(* IEC 61131-3 sources: daoli-st-library/DL_Algo (part 4) *)

(* ---- FC_DL_AccumulationZoneFillCalc.st ---- *)
(*
  DL Factory R83 | FC_DL_AccumulationZoneFillCalc
  功能：按积放区长度与料箱节距算容量件数，并算当前占位率与满料判定。
  开源溯源：无（clean-room 自研，依据公开工艺公式，来源=行业通用公式，许可证=MIT，借鉴点=公式结构）
  规则：R1-R21 全遵守
*)
FUNCTION FC_DL_AccumulationZoneFillCalc : REAL
VAR_INPUT
    fZoneLenM : REAL; // 积放区有效长度 [m] / Accumulation zone effective length [m]
    fToteLenM : REAL; // 料箱长度 [m] / Tote length [m]
    fGapMinM  : REAL; // 最小净间距 [m] / Minimum clear gap [m]
    iToteCnt  : INT;  // 区内实际料箱数 [件] / Actual totes in zone [-]
END_VAR
VAR_OUTPUT
    iCapCnt : INT;  // 区内理论容量件数 [件] / Theoretical capacity [pcs]
    fOccPct : REAL; // 占位率（实际/容量）[%] / Occupancy ratio [%]
    xFull   : BOOL; // 满料判定（占位率不低于 90%）/ Full flag, occupancy at or above 90 percent
    xValid  : BOOL; // 计算有效性标志 / Calculation validity flag
END_VAR
VAR
    fPitchM : REAL; // 单箱占用节距（箱长+净距）[m] / Per-tote pitch [m]
END_VAR
// 出口预置：四出口统一预置，满料标志预置 FALSE（安全侧）
iCapCnt := 0; fOccPct := 0.0; xFull := FALSE; xValid := FALSE;
// 非有限拦截 + 量纲自检 + 计数器域闸（R20/R21）
IF NOT (fZoneLenM > -1.0E30 AND fZoneLenM < 1.0E30) OR NOT (fToteLenM > -1.0E30 AND fToteLenM < 1.0E30) OR NOT (fGapMinM > -1.0E30 AND fGapMinM < 1.0E30) OR fZoneLenM <= 0.0 OR fToteLenM <= 0.0 OR fGapMinM < 0.0 OR iToteCnt < 0 THEN
    FC_DL_AccumulationZoneFillCalc := -1.0; RETURN; // 哨兵 -1：非有限或量纲/计数越界 / Sentinel -1
END_IF
// 单箱节距：箱长 + 最小净距，同量纲相加得 m
fPitchM := fToteLenM + fGapMinM;    // 单箱节距 [m] / Per-tote pitch [m]
// 容量：区长 ÷ 节距 向下取整（禁 TRUNC+1 写法，R28）；节距分母显式零闸（R4/R21）
IF ABS(fPitchM) > 1.0E-9 THEN       // 节距分母显式零闸 / Explicit zero gate on pitch
    iCapCnt := REAL_TO_INT(fZoneLenM / fPitchM);  // 理论容量 [件] / Theoretical capacity
ELSE
    iCapCnt := 0;                   // 除零防御缺省 [件] / Divide-by-zero default
END_IF
// 占位率：实际 ÷ 容量 × 100，容量为零时按零并标记无效（R4/R21）
IF iCapCnt > 0 THEN
    fOccPct := (INT_TO_REAL(iToteCnt) / INT_TO_REAL(iCapCnt)) * 100.0; // 占位率 [%] / Occupancy [%]
    xValid  := TRUE;                // 链路有效 / Chain valid
ELSE
    fOccPct := 0.0;                 // 容量为零不可算占位率 / Zero capacity, occupancy undefined
    xValid  := FALSE;               // 标记无效 / Flag invalid
END_IF
// 满料判定：占位率不低于 90%（含实际数超过理论容量的挤压工况）
xFull := fOccPct >= 90.0;           // 满料布尔 / Full boolean
FC_DL_AccumulationZoneFillCalc := fOccPct; // 返回占位率 [%] / Return occupancy [%]
END_FUNCTION

(* ---- FC_DL_AirDensity.st ---- *)
(*==============================================================================
 * 组件名称 (Component)  : FC_DL_AirDensity
 * 所属子库 (Sublibrary) : DL_Algo
 * 当前版本 (Version)    : 1.0.0
 * 组件分类 (Category)   : 函数（FUNCTION）· 纯函数 · 湿空气物性（密度）
 * 兼容性   (Platform)   : CODESYS 3.5 / TwinCAT 3 / 汇川 InoProShop / Schneider
 *                         Machine Expert；仅用标准 EXP / ABS / LIMIT
 * 功能描述 (Function)   : 按干空气与水蒸气分压叠加法计算湿空气密度
 *                         密度 = 干空气分压 除以 (干空气气体常数 乘以 绝对温度)
 *                                + 水蒸气分压 除以 (水蒸气气体常数 乘以 绝对温度)
 *                         单位为千克每立方米。饱和蒸汽压用 Magnus-Tetens 式计算。
 *                         用于风量质量流量换算（风机功率核算、风管风速换算）、
 *                         洁净室换气次数、烘干与涂布风量配比、空压站产气量折算。
 * 与既有件边界 (Boundary): FC_DL_HumidAirEnthalpy 出比焓（焦耳每克）；
 *                         FC_DL_DewPointCalc 出露点（摄氏度）；本件出密度
 *                         （千克每立方米）。三件共享同一 Magnus 常量口径，
 *                         但各自内联实现，禁止互相调用（泳道内零依赖），
 *                         保证任一件单独移植时不需要再带两个依赖件。
 * 精度声明 (Accuracy)   : 在零下 10 度到 50 度域内，相对误差小于 0.5 个百分点
 *                         （公开文献口径）；超出该域仅供趋势参考。这是本库对
 *                         OSCAT 同类函数行为定义的收窄，按 R11 留档。
 * 设计要点 (Key notes)  : ① 干空气分压必须防负：高湿低压的极端组态会出现
 *                           水蒸气分压大于总压，物理上不可能，但组态可给出；
 *                           出现即钳到 0 并置码，绝不输出负密度；
 *                         ② Magnus 式分母（243.12 加温度）在零下 40 度时为
 *                           203.12，恒大于 0，温度下限已保证无除零；
 *                         ③ 绝对温度由温度下限保证不小于 233.15 开，恒正；
 *                         ④ 域校验采用「钳位后继续算」策略：现场宁可要一个
 *                           标注为近似的密度值，也不要因为传感器越量程就断链。
 * 开源溯源 (Origin)     : oscat-building。参考 OSCAT 公开函数库 Building 分类
 *                         中空气密度函数的功能分类与参数域（温度 / 压力 /
 *                         湿度 三段输入，密度单值输出），只借分类、参数域与
 *                         Magnus 常量口径，实现 100% 自有 clean-room，
 *                         未复制任何源码行，不构成衍生作品。
 * 依赖     (Depends)    : 无 DL_ 内部依赖；仅 Standard.library 的 EXP 与 LIMIT
 * 故障码表 (Error codes):
 *   16#0002_1E01【信息级】温度越界被钳位
 *   16#0002_1E02【信息级】压力越界被钳位
 *   16#0002_1E03【信息级】相对湿度越界被钳位
 *   16#0002_1E04【信息级】干空气分压为负，已钳到 0（高湿低压极端组态）
 *   16#0002_1E10【信息级】入参非有限，返回 0
 * 验收向量 (Acceptance) :
 *   V1 15 度 / 101325 帕 / 湿度 0 → 约 1.2250 千克每立方米（容差 2E-3）
 *   V2 20 度 / 101325 帕 / 湿度 0 → 约 1.2041 千克每立方米（容差 2E-3）
 *   V3 20 度 / 101325 帕 / 湿度 100 → 必须小于 V2 值（水蒸气比干空气轻）
 *   V4 湿度 150 → 钳到 100，码 1E03，bValid = FALSE
 *   V5 120 度 / 50000 帕 / 湿度 100 → 触发 1E04，密度不为负
 * 红线自检 (Redline)    : R1 零全局变量表与外部变量引用 ｜ R2 零物理地址直写
 *                         R3 纯 IEC 61131-3 ｜ R4 分母恒正（温度下限保证）、
 *                         分压防负、浮点判等用容差、非有限值筛查
 *                         R5 全变量中英双语同行注释 ｜ R6 N/A（纯函数）
 *                         R7 N/A（无实例调用）
 * 修订历史 (Revision)   :
 *   2026-11-15  v1.0.0  首版入库（Round 10 · 工艺物理量链）
 *============================================================================*)

FUNCTION FC_DL_AirDensity : LREAL
VAR_INPUT
    fTempC   : LREAL := 20.0;     // 干球温度，域零下 40 到 120 [摄氏度] / Dry-bulb temperature, -40 to 120 degrees Celsius
    fPressPa : LREAL := 101325.0; // 绝对大气压，域 50000 到 120000 [帕] / Absolute pressure, 50000 to 120000 Pa
    fRh      : LREAL := 50.0;     // 相对湿度，域 0 到 100 [百分比] / Relative humidity, 0 to 100 percent
END_VAR
VAR_OUTPUT
    fDensity    : LREAL;   // 湿空气密度 [千克每立方米] / Moist air density in kilograms per cubic metre
    fSatPressPa : LREAL;   // 饱和蒸汽压，诊断与复用出口 [帕] / Saturation vapour pressure in Pa
    fVapPressPa : LREAL;   // 水蒸气分压 [帕] / Water vapour partial pressure in Pa
    bValid      : BOOL;    // 入参域全部合法且无修正事件为 TRUE [-] / TRUE when the domain is legal and no correction fired
    uErrorId    : UDINT;   // 事件码，0 = 无事件 / Event code, 0 = no event
END_VAR
VAR
    fTempUse  : LREAL;     // 生效温度（已钳位）[摄氏度] / Effective temperature
    fPressUse : LREAL;     // 生效绝对压力（已钳位）[帕] / Effective pressure
    fRhUse    : LREAL;     // 生效相对湿度（已钳位）[百分比] / Effective relative humidity
    fKelvin   : LREAL;     // 绝对温度 [开尔文] / Absolute temperature in Kelvin
    fPDry     : LREAL;     // 干空气分压 [帕] / Dry air partial pressure
    fDensDry  : LREAL;     // 干空气项密度贡献 [千克每立方米] / Dry air density contribution
    fDensVap  : LREAL;     // 水蒸气项密度贡献 [千克每立方米] / Vapour density contribution
    bDirty    : BOOL;      // 是否发生过钳位或修正事件 [-] / TRUE when any clamp or correction fired
END_VAR
VAR CONSTANT
    DL_R_DRY     : LREAL := 287.058;             // 干空气比气体常数 [焦耳每千克开] / Specific gas constant of dry air
    DL_R_VAP     : LREAL := 461.495;             // 水蒸气比气体常数 [焦耳每千克开] / Specific gas constant of water vapour
    DL_KELVIN    : LREAL := 273.15;              // 摄氏转开尔文偏移 [开] / Celsius to Kelvin offset
    DL_MAGNUS_A  : LREAL := 17.62;               // Magnus 系数 A [-] / Magnus coefficient A
    DL_MAGNUS_B  : LREAL := 243.12;              // Magnus 系数 B [摄氏度] / Magnus coefficient B
    DL_MAGNUS_C  : LREAL := 611.2;               // Magnus 基准饱和压（零度时）[帕] / Magnus reference pressure at zero Celsius
    DL_T_MIN     : LREAL := -40.0;               // 温度下限 [摄氏度] / Temperature lower bound
    DL_T_MAX     : LREAL := 120.0;               // 温度上限 [摄氏度] / Temperature upper bound
    DL_P_MIN     : LREAL := 50000.0;             // 压力下限 [帕] / Pressure lower bound
    DL_P_MAX     : LREAL := 120000.0;            // 压力上限 [帕] / Pressure upper bound
    DL_RH_MIN    : LREAL := 0.0;                 // 湿度下限 [百分比] / Humidity lower bound
    DL_RH_MAX    : LREAL := 100.0;               // 湿度上限 [百分比] / Humidity upper bound
    DL_PCT_FULL  : LREAL := 100.0;               // 百分比满量程 [-] / Full scale of the percent unit
    DL_DENS_MIN  : LREAL := 0.0;                 // 密度下限，负密度一律钳到 0 [千克每立方米] / Density lower bound
    DL_DENS_MAX  : LREAL := 20.0;                // 密度上限，覆盖高压低温极端工况 [千克每立方米] / Density upper bound
    DL_FLOAT_EPS : LREAL := 1.0E-9;              // 浮点容差 [-] / Float tolerance
    DL_BIG       : LREAL := 1.0E300;             // 非有限值兜底门限 [-] / Magnitude guard
END_VAR

(*------------------------------------------------------------------------------
 * 段 1｜输出预置
 *      Pre-set outputs
 *-----------------------------------------------------------------------------*)
FC_DL_AirDensity := 0.0;
fDensity    := 0.0;
fSatPressPa := 0.0;
fVapPressPa := 0.0;
bValid      := FALSE;
uErrorId    := 16#0000_0000;
bDirty      := FALSE;

(*------------------------------------------------------------------------------
 * 段 2｜入参有限性筛查（边界 B1）：任一非有限即返回 0 并给码
 *      Input finiteness check: any non-finite value yields zero and a code
 *-----------------------------------------------------------------------------*)
IF (fTempC <> fTempC) OR (fPressPa <> fPressPa) OR (fRh <> fRh) THEN
    uErrorId := 16#0002_1E10;
    RETURN;
END_IF

IF (ABS(fTempC) > DL_BIG) OR (ABS(fPressPa) > DL_BIG) OR (ABS(fRh) > DL_BIG) THEN
    uErrorId := 16#0002_1E10;
    RETURN;
END_IF

(*------------------------------------------------------------------------------
 * 段 3｜域校验与钳位（信息级）：钳位后继续计算，结果标注为近似
 *      Domain clamping with informational codes, computation continues
 *-----------------------------------------------------------------------------*)
fTempUse := fTempC;
IF fTempUse < DL_T_MIN THEN
    fTempUse := DL_T_MIN;
    uErrorId := 16#0002_1E01;
    bDirty   := TRUE;
ELSIF fTempUse > DL_T_MAX THEN
    fTempUse := DL_T_MAX;
    uErrorId := 16#0002_1E01;
    bDirty   := TRUE;
END_IF

fPressUse := fPressPa;
IF fPressUse < DL_P_MIN THEN
    fPressUse := DL_P_MIN;
    uErrorId  := 16#0002_1E02;
    bDirty    := TRUE;
ELSIF fPressUse > DL_P_MAX THEN
    fPressUse := DL_P_MAX;
    uErrorId  := 16#0002_1E02;
    bDirty    := TRUE;
END_IF

fRhUse := fRh;
IF fRhUse < DL_RH_MIN THEN
    fRhUse  := DL_RH_MIN;
    uErrorId := 16#0002_1E03;
    bDirty  := TRUE;
ELSIF fRhUse > DL_RH_MAX THEN
    fRhUse  := DL_RH_MAX;
    uErrorId := 16#0002_1E03;
    bDirty  := TRUE;
END_IF

(*------------------------------------------------------------------------------
 * 段 4｜饱和蒸汽压（Magnus-Tetens，单位帕）
 *      Saturation vapour pressure by the Magnus-Tetens relation in Pa
 *      分母 243.12 加温度：温度下限零下 40 度时为 203.12，恒大于 0，无除零面
 *-----------------------------------------------------------------------------*)
fSatPressPa := DL_MAGNUS_C * EXP((DL_MAGNUS_A * fTempUse) / (DL_MAGNUS_B + fTempUse));

(*------------------------------------------------------------------------------
 * 段 5｜水蒸气分压与干空气分压（防负是硬要求）
 *      Vapour partial pressure and dry air partial pressure with a negative guard
 *-----------------------------------------------------------------------------*)
fVapPressPa := fSatPressPa * (fRhUse / DL_PCT_FULL);

fPDry := fPressUse - fVapPressPa;
IF fPDry <= 0.0 THEN
    fPDry   := 0.0;              // 干空气分压不可能为负：高湿低压极端组态下的修正
    uErrorId := 16#0002_1E04;
    bDirty  := TRUE;
END_IF

(*------------------------------------------------------------------------------
 * 段 6｜绝对温度与密度叠加
 *      Absolute temperature and the density superposition
 *      fKelvin 最小为 233.15 开（由温度下限保证），恒正，无除零面
 *-----------------------------------------------------------------------------*)
fKelvin := fTempUse + DL_KELVIN;

fDensDry := fPDry / (DL_R_DRY * fKelvin);
fDensVap := fVapPressPa / (DL_R_VAP * fKelvin);
fDensity := fDensDry + fDensVap;

(*------------------------------------------------------------------------------
 * 段 7｜输出防御与有效性收口
 *      Output defence and validity close-out
 *-----------------------------------------------------------------------------*)
IF (fDensity <> fDensity) OR (ABS(fDensity) > DL_BIG) THEN
    fDensity := 0.0;             // 非有限兜底
    uErrorId := 16#0002_1E10;
    bValid   := FALSE;
    FC_DL_AirDensity := fDensity;
    RETURN;
END_IF

fDensity := LIMIT(DL_DENS_MIN, fDensity, DL_DENS_MAX);

IF bDirty THEN
    bValid := FALSE;             // 发生过钳位或修正，标注为近似
ELSE
    bValid := TRUE;
END_IF

IF ABS(fDensity) < DL_FLOAT_EPS THEN
    bValid := FALSE;             // 密度为零在物理上不可达，视为数据不可用
END_IF

FC_DL_AirDensity := fDensity;
END_FUNCTION

(* ---- FC_DL_BeltThroughputCalc.st ---- *)
(*
  DL Factory R83 | FC_DL_BeltThroughputCalc
  功能：按线速、件间距与利用率算皮带小时通过量，并给出件间净空隙。
  开源溯源：无（clean-room 自研，依据公开工艺公式，来源=行业通用公式，许可证=MIT，借鉴点=公式结构）
  规则：R1-R21 全遵守
*)
FUNCTION FC_DL_BeltThroughputCalc : REAL
VAR_INPUT
    fSpeedMps  : REAL; // 皮带线速度 [m/s] / Belt linear speed [m/s]
    fItemPitchM: REAL; // 相邻物件中心距（节距）[m] / Item pitch between centres [m]
    fItemLenM  : REAL; // 物件沿输送方向长度 [m] / Item length along travel [m]
    fUtilPct   : REAL; // 有效利用率（0~100，含停机与空载）[%] / Uptime utilisation [%]
END_VAR
VAR_OUTPUT
    fPph     : REAL; // 小时通过量 [件/h] / Throughput per hour [pcs/h]
    fGapM    : REAL; // 件间净空隙（节距-件长）[m] / Clear gap between items [m]
    fCapPps  : REAL; // 理论极限通过率（利用率 100%）[件/s] / Theoretical rate at full utilisation [pcs/s]
    xValid   : BOOL; // 计算有效性标志 / Calculation validity flag
END_VAR

// ---------- 输出预置 ----------
fPph    := 0.0;                     // 通过量清零 [件/h] / Throughput zeroed
fGapM   := 0.0;                     // 空隙清零 [m] / Gap zeroed
fCapPps := 0.0;                     // 极限率清零 [件/s] / Capability zeroed
xValid  := FALSE;                   // 有效性预置 FALSE / Validity preset FALSE

// ---------- 非有限拦截 + 量纲自检 + 节距零闸（R4/R20/R21） ----------
IF NOT (fSpeedMps > -1.0E30 AND fSpeedMps < 1.0E30) OR NOT (fItemPitchM > -1.0E30 AND fItemPitchM < 1.0E30) OR NOT (fItemLenM > -1.0E30 AND fItemLenM < 1.0E30) OR NOT (fUtilPct > -1.0E30 AND fUtilPct < 1.0E30) OR fSpeedMps <= 0.0 OR fItemPitchM <= 0.0 OR fItemLenM <= 0.0 OR fItemLenM > fItemPitchM OR fUtilPct <= 0.0 THEN
    FC_DL_BeltThroughputCalc := -1.0; // 哨兵 -1：非有限或量纲/节距越界 / Sentinel -1: non-finite or domain violation
    RETURN;
END_IF

// ---------- 利用率域闸：0~100% 之外钳位 ----------
IF fUtilPct > 100.0 THEN
    fUtilPct := 100.0;              // 上限钳位 [%] / Clamp upper bound
END_IF

// ---------- 理论极限率：m/s ÷ m = 件/s，节距分母已判正（量纲自洽） ----------
fCapPps := fSpeedMps / fItemPitchM;            // 极限通过率 [件/s] / Capability rate [pcs/s]

// ---------- 小时通过量：件/s × 3600 = 件/h，再乘利用率（含停机损失，故非恒等式） ----------
fPph := fCapPps * 3600.0 * (fUtilPct / 100.0); // 小时通过量 [件/h] / Throughput per hour [pcs/h]

// ---------- 件间净空隙：节距 - 件长，同量纲相减得 m ----------
fGapM  := fItemPitchM - fItemLenM;             // 净空隙 [m] / Clear gap [m]
xValid := TRUE;                                // 链路有效 / Chain valid
FC_DL_BeltThroughputCalc := fPph;              // 返回小时通过量 [件/h] / Return throughput [pcs/h]
END_FUNCTION

(* ---- FC_DL_BisectIterStep.st ---- *)
(* ============================================================
   DL_Algo / FC_DL_BisectIterStep ｜ v1.0.0 ｜ 2026-11-25
   功能：二分法单步。括号 [fA,fB] 取中点后按单调方向 bIncreasing 与 fFa 符号
         保留含根半区（无函数指针，故以单调性假设选定半区）
   边界：两端同号（容差判零）/ 区间退化 / 任一入参非有限 → 新括号写 0（禁 NaN/Inf
         直穿出口）、bBrktLost=TRUE（N1：判据位与实值同源，不推进）
   依赖：仅 IEC 61131-3（ABS） ｜ 溯源：DLF-B-ROOTSTEP（内部原创线）
   ============================================================ *)
FUNCTION FC_DL_BisectIterStep : BOOL
VAR_INPUT
    fA          : LREAL;  // 括号下界 [-] / Lower bracket bound
    fB          : LREAL;  // 括号上界 [-] / Upper bracket bound
    fFa         : LREAL;  // 下界函数值 [-] / Function value at the lower bound
    fFb         : LREAL;  // 上界函数值 [-] / Function value at the upper bound
    bIncreasing : BOOL;   // TRUE=f 单调递增 [-] / TRUE for a monotonically increasing residual
END_VAR
VAR_OUTPUT
    fAnew     : LREAL;  // 新括号下界 [-] / New lower bracket bound
    fBnew     : LREAL;  // 新括号上界 [-] / New upper bracket bound
    bBrktLost : BOOL;   // 括号失效或退化 [-] / Bracket lost or degenerate
END_VAR
VAR
    _fMid : LREAL;  // 中点 [-] / Midpoint of the bracket
END_VAR
VAR CONSTANT
    DL_BIS_EPS : LREAL := 1.0E-12;  // 区间退化与判零容差 [-] / Degeneracy and zero tolerance
END_VAR

(* 段 0：出口预置安全值（0，禁原始入参直穿出口，N3/R19） *)
FC_DL_BisectIterStep := FALSE;
fAnew := 0.0;  fBnew := 0.0;  bBrktLost := TRUE;

(* 段 1：非有限闸（NaN 自反 + Inf 差值自减，四入参全量枚举，R79/R272） *)
IF (fA <> fA) OR (fB <> fB) OR (fFa <> fFa) OR (fFb <> fFb) THEN RETURN; END_IF
IF ((fA - fA) <> (fA - fA)) OR ((fB - fB) <> (fB - fB))
   OR ((fFa - fFa) <> (fFa - fFa)) OR ((fFb - fFb) <> (fFb - fFb)) THEN RETURN; END_IF

(* 段 1b：闸后回传净化括号（此处起两入参已证有限，退化/同号分支可原样回传） *)
fAnew := fA;  fBnew := fB;

(* 段 1c：区间与判零闸 *)
IF ((fB - fA) - (fB - fA)) <> ((fB - fA) - (fB - fA)) THEN RETURN; END_IF
IF ABS(fB - fA) <= DL_BIS_EPS THEN RETURN; END_IF
IF (ABS(fFa) <= DL_BIS_EPS) OR (ABS(fFb) <= DL_BIS_EPS) THEN RETURN; END_IF

(* 段 2：括号有效性（fFa × fFb > 0 的同号判据，避免乘积溢出） *)
IF ((fFa > 0.0) AND (fFb > 0.0)) OR ((fFa < 0.0) AND (fFb < 0.0)) THEN RETURN; END_IF

(* 段 3：取中点并按单调方向保留含根半区 *)
_fMid := fA + (fB - fA) / 2.0;                // 中点式避免 fA+fB 溢出
IF bIncreasing THEN
    IF fFa < 0.0 THEN
        fAnew := _fMid;  fBnew := fB;         // 递增且下界为负：根在右半
    ELSE
        fAnew := fA;  fBnew := _fMid;
    END_IF
ELSE
    IF fFa < 0.0 THEN
        fAnew := fA;  fBnew := _fMid;         // 递减：半区反转
    ELSE
        fAnew := _fMid;  fBnew := fB;
    END_IF
END_IF

(* 段 4：单一出口裁决（N4） *)
bBrktLost := FALSE;  FC_DL_BisectIterStep := TRUE;
END_FUNCTION

(* ---- FC_DL_BoreCylindricityCalc.st ---- *)
(*
  DL Factory R88 | FC_DL_BoreCylindricityCalc
  功能：由两截面各四测点半径读数算圆柱度=两截面圆度取大 + 母线直线度近似，并按公差判合格
  开源溯源：无（clean-room 自研，依据公开工艺公式 圆柱度=最大圆度与母线直线度合成，许可证=MIT，借鉴点=公式结构）
  规则：R1-R16 全遵守；R88 简单件标量形（纯标量入参出参，无循环体、无方法、无属性、无数组）
*)
FUNCTION FC_DL_BoreCylindricityCalc : REAL
VAR_INPUT
    fR0Um : REAL := 50.0; // 截面 1 测点 0 半径偏差 [µm] / section 1 radius reading 0 [um]
    fR1Um : REAL := 52.0; // 截面 1 测点 1 半径偏差 [µm] / section 1 radius reading 1 [um]
    fR2Um : REAL := 49.0; // 截面 1 测点 2 半径偏差 [µm] / section 1 radius reading 2 [um]
    fR3Um : REAL := 51.0; // 截面 1 测点 3 半径偏差 [µm] / section 1 radius reading 3 [um]
    fS0Um : REAL := 53.0; // 截面 2 测点 0 半径偏差 [µm] / section 2 radius reading 0 [um]
    fS1Um : REAL := 48.0; // 截面 2 测点 1 半径偏差 [µm] / section 2 radius reading 1 [um]
    fS2Um : REAL := 55.0; // 截面 2 测点 2 半径偏差 [µm] / section 2 radius reading 2 [um]
    fS3Um : REAL := 50.0; // 截面 2 测点 3 半径偏差 [µm] / section 2 radius reading 3 [um]
    fAxisDevUm : REAL := 3.0; // 母线直线度偏差读数（轴向最大偏离） [µm] / axis straightness deviation [um]
    fTolUm : REAL := 15.0; // 圆柱度公差上限 [µm] / cylindricity tolerance [um]
END_VAR
VAR_OUTPUT
    fCylUm : REAL; // 圆柱度值（截面圆度取大 + 直线度） [µm] / cylindricity value [um]
    xPass : BOOL; // TRUE=圆柱度不超过公差 [-] / TRUE when within tolerance [-]
END_VAR
VAR
    fRound1Um : REAL; // 截面 1 圆度 [µm] / roundness of section 1 [um]
    fRound2Um : REAL; // 截面 2 圆度 [µm] / roundness of section 2 [um]
    fMaxRoundUm : REAL; // 两截面圆度取大值 [µm] / larger roundness of the two sections [um]
END_VAR

// 段 1｜出口预置
FC_DL_BoreCylindricityCalc := -1.0; // 哨兵返回 -1（无效） [-] / sentinel return -1, invalid [-]
fCylUm := 0.0; // 圆柱度预置零 [µm] / cylindricity preset zero [um]
xPass := FALSE; // 合格位预置 FALSE（未判定前不认合格） [-] / pass flag preset false [-]
fRound1Um := 0.0; // 截面 1 圆度预置零 [µm] / section 1 roundness preset zero [um]
fRound2Um := 0.0; // 截面 2 圆度预置零 [µm] / section 2 roundness preset zero [um]
fMaxRoundUm := 0.0; // 圆度大值预置零 [µm] / larger roundness preset zero [um]

// 段 2｜非有限拦截 + 域闸
IF NOT (fR0Um > -1.0E30 AND fR0Um < 1.0E30) OR NOT (fR1Um > -1.0E30 AND fR1Um < 1.0E30) OR NOT (fR2Um > -1.0E30 AND fR2Um < 1.0E30) OR NOT (fR3Um > -1.0E30 AND fR3Um < 1.0E30) THEN
    RETURN; // 截面 1 任一测点非有限即拒算 [-] / any section 1 reading non finite rejected [-]
END_IF
IF NOT (fS0Um > -1.0E30 AND fS0Um < 1.0E30) OR NOT (fS1Um > -1.0E30 AND fS1Um < 1.0E30) OR NOT (fS2Um > -1.0E30 AND fS2Um < 1.0E30) OR NOT (fS3Um > -1.0E30 AND fS3Um < 1.0E30) THEN
    RETURN; // 截面 2 任一测点非有限即拒算 [-] / any section 2 reading non finite rejected [-]
END_IF
IF NOT (fAxisDevUm > -1.0E30 AND fAxisDevUm < 1.0E30) OR NOT (fTolUm > -1.0E30 AND fTolUm < 1.0E30) THEN
    RETURN; // 直线度/公差非有限则判据静默失效，故先拦 [µm] / straightness and tolerance must be finite [um]
END_IF
IF fTolUm <= 0.0 OR fAxisDevUm < 0.0 THEN
    RETURN; // 公差正域闸 + 直线度非负闸 [µm] / positive tolerance and non negative deviation [um]
END_IF

// 段 3｜计算
fRound1Um := MAX(MAX(fR0Um, fR1Um), MAX(fR2Um, fR3Um)) - MIN(MIN(fR0Um, fR1Um), MIN(fR2Um, fR3Um)); // µm，截面 1 极差 [µm] / section 1 spread [um]
fRound2Um := MAX(MAX(fS0Um, fS1Um), MAX(fS2Um, fS3Um)) - MIN(MIN(fS0Um, fS1Um), MIN(fS2Um, fS3Um)); // µm，截面 2 极差 [µm] / section 2 spread [um]
fMaxRoundUm := MAX(fRound1Um, fRound2Um); // 两截面圆度取大 [µm] / larger of the two roundness values [um]
fCylUm := fMaxRoundUm + fAxisDevUm; // µm + µm = µm，圆柱度合成（工程近似） [µm] / [um] + [um] = [um]

// 段 4｜判定与饱和
IF NOT (fCylUm > -1.0E30 AND fCylUm < 1.0E30) THEN
    RETURN; // 结果非有限再拦一次 [-] / re-check the result for finiteness [-]
END_IF
xPass := fCylUm <= fTolUm; // 圆柱度不超过公差即合格（含边界） [µm] / within tolerance, boundary included [um]

// 段 5｜出口自检
IF fCylUm < fMaxRoundUm THEN
    RETURN; // 出口自检：合成值不得小于任一截面圆度（说明合成链被破坏） [µm] / synthetic value must not fall below [um]
END_IF
FC_DL_BoreCylindricityCalc := fCylUm; // 返回圆柱度值 [µm] / return the cylindricity value [um]
END_FUNCTION

(* ---- FC_DL_BoreRoundnessCalc.st ---- *)
(*
  DL Factory R88 | FC_DL_BoreRoundnessCalc
  功能：由固定四测点半径读数算孔圆度 (rmax-rmin)，并按 fTolUm 判合格（不用数组，逐测点标量入参）
  开源溯源：无（clean-room 自研，依据公开工艺公式 圆度最小区域近似式 R=max(r)-min(r)，许可证=MIT，借鉴点=公式结构）
  规则：R1-R16 全遵守；R88 简单件标量形（纯标量入参出参，无循环体、无方法、无属性、无数组）
*)
FUNCTION FC_DL_BoreRoundnessCalc : REAL
VAR_INPUT
    fR0Um : REAL := 50.0; // 测点 0 半径偏差读数（相对名义半径） [µm] / radius reading at point 0 [um]
    fR1Um : REAL := 52.0; // 测点 1 半径偏差读数 [µm] / radius reading at point 1 [um]
    fR2Um : REAL := 49.0; // 测点 2 半径偏差读数 [µm] / radius reading at point 2 [um]
    fR3Um : REAL := 51.0; // 测点 3 半径偏差读数 [µm] / radius reading at point 3 [um]
    fTolUm : REAL := 10.0; // 圆度公差上限 [µm] / roundness tolerance [um]
END_VAR
VAR_OUTPUT
    fRoundnessUm : REAL; // 圆度值 rmax-rmin [µm] / roundness value [um]
    xPass : BOOL; // TRUE=圆度不超过公差 [-] / TRUE when within tolerance [-]
END_VAR
VAR
    fMaxUm : REAL; // 四测点最大值 rmax [µm] / maximum radius reading [um]
    fMinUm : REAL; // 四测点最小值 rmin [µm] / minimum radius reading [um]
END_VAR

// 段 1｜出口预置
FC_DL_BoreRoundnessCalc := -1.0; // 哨兵返回 -1（无效） [-] / sentinel return -1, invalid [-]
fRoundnessUm := 0.0; // 圆度预置零 [µm] / roundness preset zero [um]
xPass := FALSE; // 合格位预置 FALSE（未判定前不认合格） [-] / pass flag preset false [-]
fMaxUm := 0.0; // 最大值预置零 [µm] / maximum preset zero [um]
fMinUm := 0.0; // 最小值预置零 [µm] / minimum preset zero [um]

// 段 2｜非有限拦截 + 域闸
IF NOT (fR0Um > -1.0E30 AND fR0Um < 1.0E30) OR NOT (fR1Um > -1.0E30 AND fR1Um < 1.0E30) THEN
    RETURN; // 测点 0/1 任一非有限即拒算 [-] / any non finite reading rejected [-]
END_IF
IF NOT (fR2Um > -1.0E30 AND fR2Um < 1.0E30) OR NOT (fR3Um > -1.0E30 AND fR3Um < 1.0E30) THEN
    RETURN; // 测点 2/3 任一非有限即拒算 [-] / any non finite reading rejected [-]
END_IF
IF NOT (fTolUm > -1.0E30 AND fTolUm < 1.0E30) THEN
    RETURN; // 公差非有限则判据静默失效，故先拦 [µm] / the tolerance must be finite [um]
END_IF
IF fTolUm <= 0.0 THEN
    RETURN; // 公差正域闸：非正公差使判定恒为不合格 [µm] / positive tolerance gate [um]
END_IF

// 段 3｜计算（四点极值法，等价 rmax-rmin 的两级 Max/Min 归约）
fMaxUm := MAX(MAX(fR0Um, fR1Um), MAX(fR2Um, fR3Um)); // 两级取大得 rmax [µm] / two stage maximum [um]
fMinUm := MIN(MIN(fR0Um, fR1Um), MIN(fR2Um, fR3Um)); // 两级取小得 rmin [µm] / two stage minimum [um]
fRoundnessUm := fMaxUm - fMinUm; // µm - µm = µm，圆度=rmax-rmin [µm] / [um] / [um] = [um]

// 段 4｜判定与饱和
IF NOT (fRoundnessUm > -1.0E30 AND fRoundnessUm < 1.0E30) THEN
    RETURN; // 结果非有限再拦一次 [-] / re-check the result for finiteness [-]
END_IF
xPass := fRoundnessUm <= fTolUm; // 圆度不超过公差即合格（含边界） [µm] / within tolerance, boundary included [um]

// 段 5｜出口自检
IF fRoundnessUm < 0.0 THEN
    RETURN; // 出口自检：圆度不得为负（负值说明极值归约出错） [µm] / roundness must not be negative [um]
END_IF
FC_DL_BoreRoundnessCalc := fRoundnessUm; // 返回圆度值 [µm] / return the roundness value [um]
END_FUNCTION

(* ---- FC_DL_BrentBracketIterStep.st ---- *)
(* ============================================================
   DL_Algo / FC_DL_BrentBracketIterStep ｜ v1.0.0 ｜ 2026-11-25
   功能：Brent 括号收缩单步（逆二次插值 + 二分混合）。三点函数值互异时按拉格朗日
         逆插值求试算点，落括号外/分母近零则退二分；由 fXLast 与 fFa 的符号关系
         收缩括号，并按宽度与 fTol 给出收敛标志
   边界：括号退化（宽度 ≤ 1E-12）→ 判已收敛；非有限 → 括号原样回传、uStepKind=0、
         bConverged=FALSE（N1）；三分母判零全用容差，禁浮点直接判等（R4）
   依赖：仅 IEC 61131-3（ABS / MIN / MAX） ｜ 溯源：DLF-B-ROOTSTEP（内部原创线）
   ============================================================ *)
FUNCTION FC_DL_BrentBracketIterStep : BOOL
VAR_INPUT
    fA      : LREAL;  // 括号下界 [-] / Lower bracket bound
    fB      : LREAL;  // 括号上界 [-] / Upper bracket bound
    fFa     : LREAL;  // 下界函数值 [-] / Function value at the lower bound
    fFb     : LREAL;  // 上界函数值 [-] / Function value at the upper bound
    fXLast  : LREAL;  // 上一步试算点 [-] / Trial point of the previous step
    fFxLast : LREAL;  // 上一步试算点函数值 [-] / Function value at the previous trial point
    fTol    : LREAL;  // 宽度收敛容差，域 > 0 [-] / Convergence tolerance on the bracket width
END_VAR
VAR_OUTPUT
    fAnew      : LREAL;  // 新括号下界 [-] / New lower bracket bound
    fBnew      : LREAL;  // 新括号上界 [-] / New upper bracket bound
    uStepKind  : UDINT;  // 步型 0 非法 / 1 逆二次插值 / 2 二分 [-] / Step kind code
    bConverged : BOOL;   // 收缩后宽度已达容差 [-] / Shrunk width within tolerance
END_VAR
VAR
    _fLo    : LREAL;  // 括号小端 [-] / Smaller bracket end
    _fHi    : LREAL;  // 括号大端 [-] / Larger bracket end
    _fMid   : LREAL;  // 二分中点 [-] / Bisection midpoint
    _fTrial : LREAL;  // 试算点 [-] / Trial point
    _fTol   : LREAL;  // 生效容差 [-] / Effective tolerance
    _bIqiOk : BOOL;   // 逆二次插值可用 [-] / Inverse quadratic interpolation usable
    _fAchk  : LREAL;  // 收缩后下界暂存 [-] / Staged lower bound
    _fBchk  : LREAL;  // 收缩后上界暂存 [-] / Staged upper bound
END_VAR
VAR CONSTANT
    DL_BRN_EPS : LREAL := 1.0E-12;  // 分母与宽度判零容差 [-] / Denominator and width tolerance
END_VAR

(* 段 0：出口预置安全侧（括号原样、步型 0、未收敛） *)
FC_DL_BrentBracketIterStep := FALSE;
fAnew := 0.0;  fBnew := 0.0;  uStepKind := 0;  bConverged := FALSE;

(* 段 1：非有限闸（七入参全量枚举，含 Inf 差值自减判） *)
IF (fA <> fA) OR (fB <> fB) OR (fFa <> fFa) OR (fFb <> fFb)
   OR (fXLast <> fXLast) OR (fFxLast <> fFxLast) OR (fTol <> fTol) THEN
    RETURN;
END_IF
IF ((fB - fA) - (fB - fA)) <> ((fB - fA) - (fB - fA)) THEN RETURN; END_IF
fAnew := fA;  fBnew := fB;                    // 闸后原样回传

(* 段 2：排序、容差兜底与退化判据 *)
_fLo := MIN(fA, fB);  _fHi := MAX(fA, fB);
IF fTol > DL_BRN_EPS THEN _fTol := fTol; ELSE _fTol := DL_BRN_EPS; END_IF
_fMid := _fLo + (_fHi - _fLo) / 2.0;
IF (_fHi - _fLo) <= DL_BRN_EPS THEN
    fAnew := _fLo;  fBnew := _fHi;  uStepKind := 2;  bConverged := TRUE;
    FC_DL_BrentBracketIterStep := TRUE;  RETURN;
END_IF

(* 段 3：逆二次插值（三分母全非零才可用，落在括号外即退二分） *)
_bIqiOk := (ABS(fFa - fFb) > DL_BRN_EPS) AND (ABS(fFa - fFxLast) > DL_BRN_EPS)
           AND (ABS(fFb - fFxLast) > DL_BRN_EPS);
_fTrial := _fMid;
IF _bIqiOk THEN
    _fTrial := fA * (fFb * fFxLast) / ((fFa - fFb) * (fFa - fFxLast))
             + fB * (fFa * fFxLast) / ((fFb - fFa) * (fFb - fFxLast))
             + fXLast * (fFa * fFb) / ((fFxLast - fFa) * (fFxLast - fFb));
    IF (_fTrial <> _fTrial) OR (_fTrial <= _fLo) OR (_fTrial >= _fHi) THEN
        _fTrial := _fMid;  _bIqiOk := FALSE;
    END_IF
END_IF

(* 段 4：括号收缩（按 fXLast 与 fFa 的符号关系取含根半区） *)
IF ((fFa > 0.0) AND (fFxLast < 0.0)) OR ((fFa < 0.0) AND (fFxLast > 0.0)) THEN
    _fAchk := MIN(fA, fXLast);  _fBchk := MAX(fA, fXLast);
ELSE
    _fAchk := MIN(fXLast, fB);  _fBchk := MAX(fXLast, fB);
END_IF

(* 段 5：无推进则退中点切分，保证迭代必推进 *)
IF (_fBchk - _fAchk) >= (_fHi - _fLo) THEN
    IF _fTrial > _fMid THEN
        _fAchk := _fMid;  _fBchk := _fHi;
    ELSE
        _fAchk := _fLo;  _fBchk := _fMid;
    END_IF
    _bIqiOk := FALSE;
END_IF

(* 段 6：单一出口裁决（N4） *)
fAnew := _fAchk;  fBnew := _fBchk;
IF _bIqiOk THEN uStepKind := 1; ELSE uStepKind := 2; END_IF
bConverged := ((_fBchk - _fAchk) <= _fTol);
IF (fAnew <> fAnew) OR (fBnew <> fBnew) THEN
    fAnew := fA;  fBnew := fB;  uStepKind := 0;  bConverged := FALSE;  RETURN;
END_IF
FC_DL_BrentBracketIterStep := TRUE;
END_FUNCTION

(* ---- FC_DL_ChkAdler32.st ---- *)
(*==============================================================================
 * 组件名称 : FC_DL_ChkAdler32 ｜ 子库 : DL_Algo ｜ v1.0.0 ｜ 2026-11-24
 * 平台     : CODESYS 3.5 / TwinCAT 3 / InoProShop / Machine Expert（纯 IEC，无厂商库）
 * 功能简介 : Adler-32 校验和（zlib / PNG 同源算法）。A 初值 1、B 初值 0，
 *            每字节 A = (A + byte) MOD 65521、B = (B + A) MOD 65521，
 *            结果 = B × 65536 + A。比 CRC 快而强度略低，适合大配方包与日志块校验。
 * 契约     : 返回 B × 65536 + A（高 16 位 B、低 16 位 A）；nLen 越界钳到 0~16；
 *            nLen = 0 时返回 1（A = 1、B = 0，空串的标准 Adler-32 值）。
 *            数组定长 ARRAY[1..16] OF BYTE（R17）。
 * 依赖     : 无 DL_ 内部依赖（R16 自足实现）；Standard.library: BYTE_TO_UDINT
 * 错误码   : R297 零码位范式：eErr 恒 0，本件结构性不置 bError
 * 红线自检 : R1 零全局 R2 零%I/%Q R3 纯IEC R4 两路累加各步取模（A<65521、B<65521），
 *            和的上界 131040 远小于 UDINT、长度先钳位后进循环 ｜ R5 双语注释
 *            R6 N/A（无状态机）R7 N/A（无定时器/沿实例）R10 标准转换
 *            R11 全声明行分号 R15 标识符零保留字冲突 R17 定长数组 R18 N/A（无 bReset）
 * 遗留假设 : 模数 65521 为小于 2^16 的最大素数（Adler 原文口径），不可换成 65535。
 * 修订历史 : 2026-11-24 R79-A 首版（校验和族 8/8）
 *============================================================================*)
FUNCTION FC_DL_ChkAdler32 : UDINT
VAR_INPUT
    aData   : ARRAY[1..16] OF BYTE;     // 待校验字节块，1..16 定长 [字节] / byte block of fixed length [byte]
    nLen    : INT;                      // 有效字节数 0~16，越界钳位 [字节] / effective length from zero to sixteen, clamped [byte]
END_VAR
VAR_OUTPUT
    eErr    : UDINT;                    // 错误码，零码位范式恒 0 / error id, always zero under the zero-code rule
    bError  : BOOL;                     // 故障标志，本件结构性不置位 / fault flag, never raised by this component
    bValid  : BOOL;                     // 结果可用标志，空块亦可用 / TRUE even for an empty block
END_VAR
VAR CONSTANT
    DL_LEN_MAX  : INT := 16;            // 字节块定长上限 [字节] / fixed block capacity [byte]
    DL_LEN_MIN  : INT := 0;             // 长度下界，0 合法 [字节] / lower length bound, zero is legal [byte]
    DL_ONE      : INT := 1;             // 数组首下标 [字节] / first array index [byte]
    DL_MOD65521 : UDINT := 65521;       // Adler 模数，小于 2^16 的最大素数 / the Adler modulus
    DL_SUM_INIT : UDINT := 1;           // A 的初值 / the initial value of the first sum
    DL_SCALE    : UDINT := 65536;       // B 的移位基数 [无量纲] / scaling factor of the second sum
    DL_ZERO_U   : UDINT := 0;           // 无符号零哨兵 / unsigned zero sentinel
END_VAR
VAR
    nSumA   : UDINT;                    // 低半累加 A，恒 < 65521 / the low half accumulator, always below the modulus
    nSumB   : UDINT;                    // 高半累加 B，恒 < 65521 / the high half accumulator, always below the modulus
    nUse    : INT;                      // 钳位后的有效长度 [字节] / effective length after clamping [byte]
    i       : INT;                      // 遍历游标 [字节] / loop cursor [byte]
END_VAR

// 段 1｜出口预置：空串的标准值为 1 / segment 1, preset the exit with the empty stream value
FC_DL_ChkAdler32 := DL_SUM_INIT;    // 缺省 1（A=1、B=0）/ default one, that is A=1 and B=0
eErr    := 0;                       // 零码位范式 / zero-code rule
bError  := FALSE;                   // 本件不产生故障级 / this component raises no fault
bValid  := TRUE;                    // 空块亦有定义 / an empty block is well defined
nSumA   := DL_SUM_INIT;             // A 初值 1 / the first sum starts at one
nSumB   := DL_ZERO_U;               // B 初值 0 / the second sum starts at zero

// 段 2｜长度钳位：越界静默整形 / segment 2, clamp the length
nUse := nLen;
IF nUse < DL_LEN_MIN THEN
    nUse := DL_LEN_MIN;             // 下越界钳到 0 / clamp to zero
ELSIF nUse > DL_LEN_MAX THEN
    nUse := DL_LEN_MAX;             // 上越界钳到定长 / clamp to the fixed capacity
END_IF

// 段 3｜两路累加：每步取模 65521，累加值恒 < 131042 不溢出 / segment 3, the two accumulators
FOR i := DL_ONE TO nUse DO
    nSumA := (nSumA + BYTE_TO_UDINT(aData[i])) MOD DL_MOD65521;     // A 累加 / accumulate the first sum
    nSumB := (nSumB + nSumA) MOD DL_MOD65521;                       // B 累加 A / accumulate the second sum over the first
END_FOR

// 段 4｜出口：B 在高半、A 在低半 / segment 4, exit with B in the high half
FC_DL_ChkAdler32 := (nSumB * DL_SCALE) + nSumA;
END_FUNCTION

(* ---- FC_DL_ChkFletcher16.st ---- *)
(*==============================================================================
 * 组件名称 : FC_DL_ChkFletcher16 ｜ 子库 : DL_Algo ｜ v1.0.0 ｜ 2026-11-24
 * 平台     : CODESYS 3.5 / TwinCAT 3 / InoProShop / Machine Expert（纯 IEC，无厂商库）
 * 功能简介 : 标准 Fletcher-16 校验和。两路累加：sum1 逐字节累加、sum2 累加 sum1，
 *            二者每步各取模 255，结果 = sum2 × 256 + sum1。相比简单字节和，
 *            Fletcher 对字节换位与丢字节敏感，适合串口帧、条码回读、配方块校验。
 * 契约     : 返回 32 位结果（高 16 位 sum2、低 16 位 sum1，各 < 255）；
 *            nLen 越界钳到 0~16（钳位不报错，属输入整形）；nLen = 0 返回 0。
 *            数组定长 ARRAY[1..16] OF BYTE（R17）。
 * 依赖     : 无 DL_ 内部依赖（R16 自足实现）；Standard.library: BYTE_TO_UDINT
 * 错误码   : R297 零码位范式：eErr 恒 0，本件结构性不置 bError
 * 红线自检 : R1 零全局 R2 零%I/%Q R3 纯IEC R4 长度先钳位后进循环、取模除数恒为常量 255、
 *            累加上界 255+254 不溢出 ｜ R5 双语注释 R6 N/A（无状态机）
 *            R7 N/A（无定时器/沿实例）R10 标准转换 R11 全声明行分号
 *            R15 标识符零保留字冲突 R17 定长数组 R18 N/A（无 bReset）
 * 遗留假设 : 模数取 255（Fletcher 原始口径，非 256）；与某些实现的 255 vs 256 差异
 *            会导致校验不一致，对接第三方协议前须核对其模数口径。
 * 修订历史 : 2026-11-24 R79-A 首版（校验和族 1/8）
 *============================================================================*)
FUNCTION FC_DL_ChkFletcher16 : UDINT
VAR_INPUT
    aData   : ARRAY[1..16] OF BYTE;     // 待校验字节块，1..16 定长 [字节] / byte block of fixed length [byte]
    nLen    : INT;                      // 有效字节数 0~16，越界钳位 [字节] / effective length from zero to sixteen, clamped [byte]
END_VAR
VAR_OUTPUT
    eErr    : UDINT;                    // 错误码，零码位范式恒 0 / error id, always zero under the zero-code rule
    bError  : BOOL;                     // 故障标志，本件结构性不置位 / fault flag, never raised by this component
    bValid  : BOOL;                     // 结果可用标志，空块亦可用 / TRUE even for an empty block
END_VAR
VAR CONSTANT
    DL_LEN_MAX : INT := 16;             // 字节块定长上限 [字节] / fixed block capacity [byte]
    DL_LEN_MIN : INT := 0;              // 长度下界，0 合法 [字节] / lower length bound, zero is legal [byte]
    DL_ONE     : INT := 1;              // 数组首下标 [字节] / first array index [byte]
    DL_MOD255  : UDINT := 255;          // Fletcher 模数 [无量纲] / the Fletcher modulus
    DL_SCALE   : UDINT := 256;          // 高字节移位基数 [无量纲] / high byte scaling factor
    DL_ZERO_U  : UDINT := 0;            // 无符号零哨兵 / unsigned zero sentinel
END_VAR
VAR
    nSum1   : UDINT;                    // 字节累加和 [无量纲] / running byte sum
    nSum2   : UDINT;                    // sum1 的累加和 [无量纲] / running sum of the first sum
    nUse    : INT;                      // 钳位后的有效长度 [字节] / effective length after clamping [byte]
    i       : INT;                      // 遍历游标 [字节] / loop cursor [byte]
END_VAR

// 段 1｜出口预置 / segment 1, preset the exit
FC_DL_ChkFletcher16 := DL_ZERO_U;   // 缺省 0 / default zero
eErr   := 0;                        // 零码位范式 / zero-code rule
bError := FALSE;                    // 本件不产生故障级 / this component raises no fault
bValid := TRUE;                     // 空块亦有定义，结果恒可用 / an empty block is well defined
nSum1  := DL_ZERO_U;                // 第一路累加器清零 / clear the first accumulator
nSum2  := DL_ZERO_U;                // 第二路累加器清零 / clear the second accumulator

// 段 2｜长度钳位：越界静默整形，不进故障态 / segment 2, clamp the length
nUse := nLen;
IF nUse < DL_LEN_MIN THEN
    nUse := DL_LEN_MIN;             // 下越界钳到 0 / clamp to zero
ELSIF nUse > DL_LEN_MAX THEN
    nUse := DL_LEN_MAX;             // 上越界钳到定长 / clamp to the fixed capacity
END_IF

// 段 3｜两路累加：每步取模 255，累加值恒 < 255 故不会溢出 / segment 3, the two accumulators
FOR i := DL_ONE TO nUse DO
    nSum1 := (nSum1 + BYTE_TO_UDINT(aData[i])) MOD DL_MOD255;   // 字节和 / byte sum
    nSum2 := (nSum2 + nSum1) MOD DL_MOD255;                     // 字节和的累加 / sum of the sums
END_FOR

// 段 4｜出口：高半 sum2、低半 sum1 / segment 4, exit with sum two in the high half
FC_DL_ChkFletcher16 := (nSum2 * DL_SCALE) + nSum1;
END_FUNCTION

(* ---- FC_DL_ChkFletcher32.st ---- *)
(*==============================================================================
 * 组件名称 : FC_DL_ChkFletcher32 ｜ 子库 : DL_Algo ｜ v1.0.0 ｜ 2026-11-24
 * 平台     : CODESYS 3.5 / TwinCAT 3 / InoProShop / Machine Expert（纯 IEC，无厂商库）
 * 功能简介 : Fletcher-32 校验和 —— 把字节流按 16 位小端字处理，两路累加各取模 65535，
 *            结果 = sum2 × 65536 + sum1。奇数长度时末字节作低字节、高字节补零成字
 *            （与「末字节补零」的通行口径一致）。用于长帧（>512 字节）与文件块校验。
 * 契约     : 返回 32 位结果；nLen 越界钳到 0~16；nLen = 0 返回 0。
 *            数组定长 ARRAY[1..16] OF BYTE（R17）。
 * 依赖     : 无 DL_ 内部依赖（R16 自足实现）；Standard.library: BYTE_TO_UDINT
 * 错误码   : R297 零码位范式：eErr 恒 0，本件结构性不置 bError
 * 红线自检 : R1 零全局 R2 零%I/%Q R3 纯IEC R4 字下标经上界复核（2k ≤ nUse 才取高字节）、
 *            累加上界 65535+65534 < 2^32、取模除数恒为常量 ｜ R5 双语注释
 *            R6 N/A（无状态机）R7 N/A（无定时器/沿实例）R10 标准转换
 *            R11 全声明行分号 R15 标识符零保留字冲突 R17 定长数组 R18 N/A（无 bReset）
 * 遗留假设 : 小端组装（低字节在前）；大端协议须调用方先换序，本件不做字节序猜测。
 * 修订历史 : 2026-11-24 R79-A 首版（校验和族 2/8）
 *============================================================================*)
FUNCTION FC_DL_ChkFletcher32 : UDINT
VAR_INPUT
    aData   : ARRAY[1..16] OF BYTE;     // 待校验字节块，1..16 定长 [字节] / byte block of fixed length [byte]
    nLen    : INT;                      // 有效字节数 0~16，越界钳位 [字节] / effective length from zero to sixteen, clamped [byte]
END_VAR
VAR_OUTPUT
    eErr    : UDINT;                    // 错误码，零码位范式恒 0 / error id, always zero under the zero-code rule
    bError  : BOOL;                     // 故障标志，本件结构性不置位 / fault flag, never raised by this component
    bValid  : BOOL;                     // 结果可用标志，空块亦可用 / TRUE even for an empty block
END_VAR
VAR CONSTANT
    DL_LEN_MAX : INT := 16;             // 字节块定长上限 [字节] / fixed block capacity [byte]
    DL_LEN_MIN : INT := 0;              // 长度下界，0 合法 [字节] / lower length bound, zero is legal [byte]
    DL_ONE     : INT := 1;              // 数组首下标 [字节] / first array index [byte]
    DL_TWO     : INT := 2;              // 每字字节数与奇偶判断基数 [字节] / bytes per word and the parity radix [byte]
    DL_MOD16   : UDINT := 65535;        // Fletcher-32 模数 [无量纲] / the Fletcher thirty two modulus
    DL_SCALE   : UDINT := 65536;        // 高半字移位基数 [无量纲] / high word scaling factor
    DL_BYTE_SH : UDINT := 256;          // 字节移位基数 [无量纲] / byte scaling factor
    DL_ZERO_U  : UDINT := 0;            // 无符号零哨兵 / unsigned zero sentinel
END_VAR
VAR
    nSum1   : UDINT;                    // 字累加和 [无量纲] / running word sum
    nSum2   : UDINT;                    // sum1 的累加和 [无量纲] / running sum of the first sum
    nWord   : UDINT;                    // 当前 16 位小端字 [无量纲] / the current little endian word
    nLo     : UDINT;                    // 字内低字节 [无量纲] / low byte of the word
    nHi     : UDINT;                    // 字内高字节，奇数长度时为 0 [无量纲] / high byte, zero on an odd tail
    nUse    : INT;                      // 钳位后的有效长度 [字节] / effective length after clamping [byte]
    nWords  : INT;                      // 字数，奇数长度向上取整 [字] / word count rounded up [word]
    k       : INT;                      // 字游标 [字] / word cursor [word]
    nIdx    : INT;                      // 字内第二个字节的数组下标 [字节] / index of the second byte in the word [byte]
END_VAR

// 段 1｜出口预置 / segment 1, preset the exit
FC_DL_ChkFletcher32 := DL_ZERO_U;   // 缺省 0 / default zero
eErr   := 0;                        // 零码位范式 / zero-code rule
bError := FALSE;                    // 本件不产生故障级 / this component raises no fault
bValid := TRUE;                     // 空块亦有定义 / an empty block is well defined
nSum1  := DL_ZERO_U;                // 第一路累加器清零 / clear the first accumulator
nSum2  := DL_ZERO_U;                // 第二路累加器清零 / clear the second accumulator

// 段 2｜长度钳位与字数换算：奇数长度向上取整成字 / segment 2, clamp the length and round the word count up
nUse := nLen;
IF nUse < DL_LEN_MIN THEN
    nUse := DL_LEN_MIN;             // 下越界钳到 0 / clamp to zero
ELSIF nUse > DL_LEN_MAX THEN
    nUse := DL_LEN_MAX;             // 上越界钳到定长 / clamp to the fixed capacity
END_IF
nWords := (nUse + DL_ONE) / DL_TWO; // 向上取整的字数 / the word count rounded up

// 段 3｜逐字累加：低字节在前，奇数尾字节高半补零 / segment 3, word by word with a zero padded tail
FOR k := DL_ONE TO nWords DO
    nLo  := BYTE_TO_UDINT(aData[(DL_TWO * k) - DL_ONE]);    // 低字节，下标必 ≤ nUse / the low byte, its index never exceeds the length
    nHi  := DL_ZERO_U;                                      // 高字节缺省 0，即补零成字 / the high byte defaults to zero, padding the word
    nIdx := DL_TWO * k;                                     // 高字节下标 / the index of the high byte
    IF nIdx <= nUse THEN
        nHi := BYTE_TO_UDINT(aData[nIdx]);                   // 长度允许才取高字节 / take the high byte only when the length allows
    END_IF
    nWord := nLo + (nHi * DL_BYTE_SH);                       // 小端组装 / little endian assembly
    nSum1 := (nSum1 + nWord) MOD DL_MOD16;                   // 字和 / word sum
    nSum2 := (nSum2 + nSum1) MOD DL_MOD16;                   // 字和的累加 / sum of the sums
END_FOR

// 段 4｜出口：高半 sum2、低半 sum1 / segment 4, exit with sum two in the high half
FC_DL_ChkFletcher32 := (nSum2 * DL_SCALE) + nSum1;
END_FUNCTION

(* ---- FC_DL_ChkParityBlock.st ---- *)
(*==============================================================================
 * 组件名称 : FC_DL_ChkParityBlock ｜ 子库 : DL_Algo ｜ v1.0.0 ｜ 2026-11-24
 * 平台     : CODESYS 3.5 / TwinCAT 3 / InoProShop / Machine Expert（纯 IEC，无厂商库）
 * 功能简介 : 整块字节的偶校验结论。统计全块为 1 的比特总数，总数为偶数返回 TRUE。
 *            与逐帧奇偶校验位同源：发送端把本件结果放进校验位，接收端对「数据 + 校验位」
 *            复算应得 FALSE（偶数个 1）。用于老式 ASCII 链路、条码枪回读的一致性核验。
 * 契约     : 返回 TRUE 表示 1 的个数为偶数（偶校验成立）；nLen 越界钳到 0~16；
 *            nLen = 0 时 1 的个数为 0（偶数），返回 TRUE。
 *            数组定长 ARRAY[1..16] OF BYTE（R17）。
 * 依赖     : 无 DL_ 内部依赖（R16 自足实现）；Standard.library: BYTE_TO_UDINT
 * 错误码   : R297 零码位范式：eErr 恒 0，本件结构性不置 bError
 * 红线自检 : R1 零全局 R2 零%I/%Q R3 纯IEC R4 位计数用整除取余循环（每字节最多 8 次）、
 *            长度先钳位后进循环 ｜ R5 双语注释 R6 N/A（无状态机）
 *            R7 N/A（无定时器/沿实例）R10 标准转换 R11 全声明行分号
 *            R15 标识符零保留字冲突 R17 定长数组 R18 N/A（无 bReset）
 * 遗留假设 : 「偶校验」定义为整块比特和为偶数；若协议要求「校验位使总数成偶」，
 *            则须在接收侧把校验位一并送入本件，判据取 FALSE。
 * 修订历史 : 2026-11-24 R79-A 首版（校验和族 7/8）
 *============================================================================*)
FUNCTION FC_DL_ChkParityBlock : BOOL
VAR_INPUT
    aData   : ARRAY[1..16] OF BYTE;     // 待校验字节块，1..16 定长 [字节] / byte block of fixed length [byte]
    nLen    : INT;                      // 有效字节数 0~16，越界钳位 [字节] / effective length from zero to sixteen, clamped [byte]
END_VAR
VAR_OUTPUT
    eErr    : UDINT;                    // 错误码，零码位范式恒 0 / error id, always zero under the zero-code rule
    bError  : BOOL;                     // 故障标志，本件结构性不置位 / fault flag, never raised by this component
    bValid  : BOOL;                     // 结果可用标志，空块亦可用 / TRUE even for an empty block
    nBitOnes : UDINT;                   // 整块为 1 的比特总数，供诊断 / total number of one bits, for diagnostics
END_VAR
VAR CONSTANT
    DL_LEN_MAX : INT := 16;             // 字节块定长上限 [字节] / fixed block capacity [byte]
    DL_LEN_MIN : INT := 0;              // 长度下界，0 合法 [字节] / lower length bound, zero is legal [byte]
    DL_ONE     : INT := 1;              // 数组首下标 [字节] / first array index [byte]
    DL_TWO     : UDINT := 2;            // 位提取的进制基数 [无量纲] / radix of the bit extraction
    DL_EVEN    : UDINT := 2;            // 奇偶判断的模数 [无量纲] / modulus of the parity test
    DL_ZERO_U  : UDINT := 0;            // 无符号零哨兵 / unsigned zero sentinel
END_VAR
VAR
    nByte   : UDINT;                    // 当前字节的位提取工作副本 / working copy of the current byte
    nOnes   : UDINT;                    // 累计的 1 比特数 / accumulated one bits
    nUse    : INT;                      // 钳位后的有效长度 [字节] / effective length after clamping [byte]
    i       : INT;                      // 遍历游标 [字节] / loop cursor [byte]
END_VAR

// 段 1｜出口预置 / segment 1, preset the exit
FC_DL_ChkParityBlock := TRUE;       // 缺省偶校验成立（零个 1）/ default even parity, zero one bits
eErr     := 0;                      // 零码位范式 / zero-code rule
bError   := FALSE;                  // 本件不产生故障级 / this component raises no fault
bValid   := TRUE;                   // 空块亦有定义 / an empty block is well defined
nOnes    := DL_ZERO_U;              // 比特计数清零 / clear the bit counter
nBitOnes := DL_ZERO_U;              // 诊断出口清零 / clear the diagnostic output

// 段 2｜长度钳位：越界静默整形 / segment 2, clamp the length
nUse := nLen;
IF nUse < DL_LEN_MIN THEN
    nUse := DL_LEN_MIN;             // 下越界钳到 0 / clamp to zero
ELSIF nUse > DL_LEN_MAX THEN
    nUse := DL_LEN_MAX;             // 上越界钳到定长 / clamp to the fixed capacity
END_IF

// 段 3｜逐字节取位计数：右移一位即整除 2，最低位即取余 / segment 3, count the one bits byte by byte
FOR i := DL_ONE TO nUse DO
    nByte := BYTE_TO_UDINT(aData[i]);   // 取当前字节 / take the current byte
    WHILE nByte > DL_ZERO_U DO
        nOnes := nOnes + (nByte MOD DL_TWO);    // 最低位为 1 则加一 / add one when the low bit is set
        nByte := nByte / DL_TWO;                // 右移一位 / shift one bit right
    END_WHILE
END_FOR

// 段 4｜出口：总数为偶数即偶校验成立 / segment 4, even parity holds when the total is even
nBitOnes := nOnes;                              // 诊断出口 / the diagnostic output
FC_DL_ChkParityBlock := ((nOnes MOD DL_EVEN) = DL_ZERO_U);
END_FUNCTION

(* ---- FC_DL_ChkSum32Mod.st ---- *)
(*==============================================================================
 * 组件名称 : FC_DL_ChkSum32Mod ｜ 子库 : DL_Algo ｜ v1.0.0 ｜ 2026-11-24
 * 平台     : CODESYS 3.5 / TwinCAT 3 / InoProShop / Machine Expert（纯 IEC，无厂商库）
 * 功能简介 : 32 位字求和取模校验。字节流按 4 字节小端组装成 32 位字累加，
 *            最后返回 sum MOD 16#FFFF_FFFF。文件块、固件包、大配方块的轻量完整性校验。
 *            实现要点：不先做「四字组装再求和」——那样最多 4×16#FFFF_FFFF 会溢出 UDINT；
 *            改为按字节加权（权 1/256/65536/16777216 循环）并用「减模数」法逐步归一，
 *            nAcc 恒 < 16#FFFF_FFFF，任何一步都不溢出。尾字节不足 4 个即权值循环自然补零。
 * 契约     : 返回 sum MOD 16#FFFF_FFFF（0~16#FFFF_FFFE）；nLen 越界钳到 0~16；nLen = 0 返回 0。
 *            数组定长 ARRAY[1..16] OF BYTE（R17）。
 * 依赖     : 无 DL_ 内部依赖（R16 自足实现）；Standard.library: BYTE_TO_UDINT
 * 错误码   : R297 零码位范式：eErr 恒 0，本件结构性不置 bError
 * 红线自检 : R1 零全局 R2 零%I/%Q R3 纯IEC R4 单项 ≤ 255×2^24 < 模数故累加一次归一即足、
 *            权值乘前先判上界防回绕、NOT 用位反 ｜ R5 双语注释 R6 N/A（无状态机）
 *            R7 N/A（无定时器/沿实例）R10 标准转换 R11 全声明行分号
 *            R15 标识符零保留字冲突 R17 定长数组 R18 N/A（无 bReset）
 * 遗留假设 : 小端组装；「sum MOD 16#FFFF_FFFF」为协议原始口径（不是 2^32 回绕），
 *            两者在第 16#FFFF_FFFF 个字节才分岔，本件按协议原文实现。
 * 修订历史 : 2026-11-24 R79-A 首版（校验和族 6/8）
 *============================================================================*)
FUNCTION FC_DL_ChkSum32Mod : UDINT
VAR_INPUT
    aData   : ARRAY[1..16] OF BYTE;     // 待校验字节块，1..16 定长 [字节] / byte block of fixed length [byte]
    nLen    : INT;                      // 有效字节数 0~16，越界钳位 [字节] / effective length from zero to sixteen, clamped [byte]
END_VAR
VAR_OUTPUT
    eErr    : UDINT;                    // 错误码，零码位范式恒 0 / error id, always zero under the zero-code rule
    bError  : BOOL;                     // 故障标志，本件结构性不置位 / fault flag, never raised by this component
    bValid  : BOOL;                     // 结果可用标志，空块亦可用 / TRUE even for an empty block
END_VAR
VAR CONSTANT
    DL_LEN_MAX  : INT := 16;            // 字节块定长上限 [字节] / fixed block capacity [byte]
    DL_LEN_MIN  : INT := 0;             // 长度下界，0 合法 [字节] / lower length bound, zero is legal [byte]
    DL_ONE      : INT := 1;             // 数组首下标 [字节] / first array index [byte]
    DL_MOD_MASK : UDINT := 16#FFFF_FFFF;    // 取模的模数 [无量纲] / the modulus of the protocol
    DL_SHIFT_MAX : UDINT := 16#0100_0000;   // 最高字节权 2^24，再乘 256 会回绕 [无量纲] / the top byte weight, the next step would wrap
    DL_ONE_U    : UDINT := 1;           // 无符号一，权值循环起点 [无量纲] / unsigned one, the first weight
    DL_BYTE_SH  : UDINT := 256;         // 字节权倍数 [无量纲] / weight multiplier per byte
    DL_ZERO_U   : UDINT := 0;           // 无符号零哨兵 / unsigned zero sentinel
END_VAR
VAR
    nAcc    : UDINT;                    // 逐步归一的累加器，恒 < 模数 / the reduced accumulator, always below the modulus
    nTerm   : UDINT;                    // 当前字节的加权项，最大 255×2^24 / the weighted term of one byte
    nShift  : UDINT;                    // 当前字节权 1/256/65536/16777216 循环 [无量纲] / the weight cycling over four bytes
    nUse    : INT;                      // 钳位后的有效长度 [字节] / effective length after clamping [byte]
    i       : INT;                      // 遍历游标 [字节] / loop cursor [byte]
END_VAR

// 段 1｜出口预置 / segment 1, preset the exit
FC_DL_ChkSum32Mod := DL_ZERO_U;
eErr    := 0;                       // 零码位范式 / zero-code rule
bError  := FALSE;                   // 本件不产生故障级 / this component raises no fault
bValid  := TRUE;                    // 空块亦有定义 / an empty block is well defined
nAcc    := DL_ZERO_U;               // 累加器清零 / clear the accumulator
nShift  := DL_ONE_U;                // 首字节权为 1 / the first byte weighs one

// 段 2｜长度钳位：越界静默整形 / segment 2, clamp the length
nUse := nLen;
IF nUse < DL_LEN_MIN THEN
    nUse := DL_LEN_MIN;             // 下越界钳到 0 / clamp to zero
ELSIF nUse > DL_LEN_MAX THEN
    nUse := DL_LEN_MAX;             // 上越界钳到定长 / clamp to the fixed capacity
END_IF

// 段 3｜逐字节加权并减模数归一：单项必小于模数，故一次减法即够 / segment 3, weighted accumulation with a single reduction
FOR i := DL_ONE TO nUse DO
    nTerm := BYTE_TO_UDINT(aData[i]) * nShift;      // 加权项 ≤ 255×2^24 = 16#FF00_0000，远小于模数 / the term stays well below the modulus
    IF nAcc >= (DL_MOD_MASK - nTerm) THEN
        nAcc := nAcc - (DL_MOD_MASK - nTerm);       // 等价于 nAcc + nTerm − 模数，且不产生中间溢出 / equals the sum minus the modulus
    ELSE
        nAcc := nAcc + nTerm;                       // 未越模数直接加上 / plain accumulation when no reduction is needed
    END_IF
    IF nShift = DL_SHIFT_MAX THEN
        nShift := DL_ONE_U;                         // 第 5 个字节权回到 1，相当于补齐成 4 字节字 / the fifth byte restarts the word
    ELSE
        nShift := nShift * DL_BYTE_SH;              // 乘前已判上界，不会回绕 / the bound was checked, no wrap
    END_IF
END_FOR

// 段 4｜出口：累加器已归一到 [0, 模数) / segment 4, exit with a reduced accumulator
FC_DL_ChkSum32Mod := nAcc;
END_FUNCTION

(* ---- FC_DL_ChkTwosCompSum16.st ---- *)
(*==============================================================================
 * 组件名称 : FC_DL_ChkTwosCompSum16 ｜ 子库 : DL_Algo ｜ v1.0.0 ｜ 2026-11-24
 * 平台     : CODESYS 3.5 / TwinCAT 3 / InoProShop / Machine Expert（纯 IEC，无厂商库）
 * 功能简介 : 16 位字求和二补数校验（two's complement checksum，串口协议常用的
 *            「求和取反加一」帧尾）。字节流按 16 位小端字累加，再取 16#10000 − (sum MOD
 *            16#10000)；结果落在 16#0001~16#FFFF，0 用原码 0 表示（不进位到 16#10000）。
 * 契约     : 返回二补数校验值（0~16#FFFF）；nLen 越界钳到 0~16；nLen = 0 返回 0。
 *            奇数长度时末字节作低字节、高字节补零。
 *            数组定长 ARRAY[1..16] OF BYTE（R17）。
 * 依赖     : 无 DL_ 内部依赖（R16 自足实现）；Standard.library: BYTE_TO_UDINT
 * 错误码   : R297 零码位范式：eErr 恒 0，本件结构性不置 bError
 * 红线自检 : R1 零全局 R2 零%I/%Q R3 纯IEC R4 字下标经上界复核、累加上界 8×65535 不溢出、
 *            补码零特判（16#10000 不可表示） ｜ R5 双语注释 R6 N/A（无状态机）
 *            R7 N/A（无定时器/沿实例）R10 标准转换 R11 全声明行分号
 *            R15 标识符零保留字冲突 R17 定长数组 R18 N/A（无 bReset）
 * 遗留假设 : 小端组装；某些协议口径为「大端字序」或「字节和取补」，对接前须核对协议原文。
 * 修订历史 : 2026-11-24 R79-A 首版（校验和族 5/8）
 *============================================================================*)
FUNCTION FC_DL_ChkTwosCompSum16 : UDINT
VAR_INPUT
    aData   : ARRAY[1..16] OF BYTE;     // 待校验字节块，1..16 定长 [字节] / byte block of fixed length [byte]
    nLen    : INT;                      // 有效字节数 0~16，越界钳位 [字节] / effective length from zero to sixteen, clamped [byte]
END_VAR
VAR_OUTPUT
    eErr    : UDINT;                    // 错误码，零码位范式恒 0 / error id, always zero under the zero-code rule
    bError  : BOOL;                     // 故障标志，本件结构性不置位 / fault flag, never raised by this component
    bValid  : BOOL;                     // 结果可用标志，空块亦可用 / TRUE even for an empty block
END_VAR
VAR CONSTANT
    DL_LEN_MAX  : INT := 16;            // 字节块定长上限 [字节] / fixed block capacity [byte]
    DL_LEN_MIN  : INT := 0;             // 长度下界，0 合法 [字节] / lower length bound, zero is legal [byte]
    DL_ONE      : INT := 1;             // 数组首下标 [字节] / first array index [byte]
    DL_TWO      : INT := 2;             // 每字字节数与奇偶基数 [字节] / bytes per word and the parity radix [byte]
    DL_WORD_MOD : UDINT := 65536;       // 16 位字回绕基数 [无量纲] / the sixteen bit wrap modulus
    DL_BYTE_SH  : UDINT := 256;         // 字节移位基数 [无量纲] / byte scaling factor
    DL_ZERO_U   : UDINT := 0;           // 无符号零哨兵 / unsigned zero sentinel
END_VAR
VAR
    nSum    : UDINT;                    // 字累加和，最大 8×65535 远小于上界 / word sum, at most eight times sixty five thousand
    nWord   : UDINT;                    // 当前 16 位小端字 [无量纲] / the current little endian word
    nLo     : UDINT;                    // 字内低字节 [无量纲] / low byte of the word
    nHi     : UDINT;                    // 字内高字节，奇数长度时为 0 [无量纲] / high byte, zero on an odd tail
    nLow16  : UDINT;                    // 累加和的低 16 位 [无量纲] / the low sixteen bits of the sum
    nUse    : INT;                      // 钳位后的有效长度 [字节] / effective length after clamping [byte]
    nWords  : INT;                      // 字数，奇数长度向上取整 [字] / word count rounded up [word]
    k       : INT;                      // 字游标 [字] / word cursor [word]
    nIdx    : INT;                      // 字内第二个字节的下标 [字节] / index of the second byte in the word [byte]
END_VAR

// 段 1｜出口预置 / segment 1, preset the exit
FC_DL_ChkTwosCompSum16 := DL_ZERO_U;
eErr   := 0;                        // 零码位范式 / zero-code rule
bError := FALSE;                    // 本件不产生故障级 / this component raises no fault
bValid := TRUE;                     // 空块亦有定义 / an empty block is well defined
nSum   := DL_ZERO_U;                // 累加器清零 / clear the accumulator

// 段 2｜长度钳位与字数换算 / segment 2, clamp the length and round the word count up
nUse := nLen;
IF nUse < DL_LEN_MIN THEN
    nUse := DL_LEN_MIN;             // 下越界钳到 0 / clamp to zero
ELSIF nUse > DL_LEN_MAX THEN
    nUse := DL_LEN_MAX;             // 上越界钳到定长 / clamp to the fixed capacity
END_IF
nWords := (nUse + DL_ONE) / DL_TWO;

// 段 3｜逐字累加：低字节在前，尾字节高半补零 / segment 3, word by word with a zero padded tail
FOR k := DL_ONE TO nWords DO
    nLo  := BYTE_TO_UDINT(aData[(DL_TWO * k) - DL_ONE]);    // 低字节，下标必 ≤ nUse / the low byte, always inside the block
    nHi  := DL_ZERO_U;                                      // 补零缺省 / padding default
    nIdx := DL_TWO * k;                                     // 高字节下标 / the high byte index
    IF nIdx <= nUse THEN
        nHi := BYTE_TO_UDINT(aData[nIdx]);                   // 长度允许才取 / taken only when the length allows
    END_IF
    nWord := nLo + (nHi * DL_BYTE_SH);                       // 小端组装 / little endian assembly
    nSum  := nSum + nWord;                                   // 宽域累加，无回绕 / wide accumulation without wrap
END_FOR

// 段 4｜二补数：低 16 位取反加一；为 0 时用原码 0 表示 / segment 4, the two's complement
nLow16 := nSum MOD DL_WORD_MOD;         // 低 16 位 / the low sixteen bits
IF nLow16 = DL_ZERO_U THEN
    FC_DL_ChkTwosCompSum16 := DL_ZERO_U;    // 补码会得 16#10000，不可表示，用 0 表示 / the complement would be sixteen to the fourth, use zero
ELSE
    FC_DL_ChkTwosCompSum16 := DL_WORD_MOD - nLow16;
END_IF
END_FUNCTION

(* ---- FC_DL_ChuteFullPredict.st ---- *)
(*
  DL Factory R83 | FC_DL_ChuteFullPredict
  功能：按入流与出流净流量预测滑槽从当前填充率到满料所需时间。
  开源溯源：无（clean-room 自研，依据公开工艺公式，来源=行业通用公式，许可证=MIT，借鉴点=公式结构）
  规则：R1-R21 全遵守
*)
FUNCTION FC_DL_ChuteFullPredict : REAL
VAR_INPUT
    fFillPct     : REAL; // 当前填充率（0~100）[%] / Current fill ratio [%]
    fInflowPpm   : REAL; // 入流件率 [件/min] / Inflow rate [pcs/min]
    fOutflowPpm  : REAL; // 出流件率 [件/min] / Outflow rate [pcs/min]
    fCapacityPcs : REAL; // 滑槽容量 [件] / Chute capacity [pcs]
END_VAR
VAR_OUTPUT
    fNetPpm      : REAL; // 净流入件率（入-出）[件/min] / Net accumulation rate [pcs/min]
    fTimeToFullS : REAL; // 到满料剩余时间（净流非正时为 0）[s] / Time to full, 0 = never [s]
    xCritical    : BOOL; // 满料风险（净流入且剩余不足 60 s）/ Full-risk flag
    xValid       : BOOL; // 计算有效性标志 / Calculation validity flag
END_VAR
VAR
    fRoomPcs : REAL; // 剩余可容纳件数 [件] / Remaining free capacity [pcs]
END_VAR
fNetPpm := 0.0; fTimeToFullS := 0.0; xCritical := FALSE; xValid := FALSE;  // 出口预置（安全侧）
// 非有限拦截 + 量纲自检（R20/R21）
IF NOT (fFillPct > -1.0E30 AND fFillPct < 1.0E30) OR NOT (fInflowPpm > -1.0E30 AND fInflowPpm < 1.0E30) OR NOT (fOutflowPpm > -1.0E30 AND fOutflowPpm < 1.0E30) OR NOT (fCapacityPcs > -1.0E30 AND fCapacityPcs < 1.0E30) OR fInflowPpm < 0.0 OR fOutflowPpm < 0.0 OR fCapacityPcs <= 0.0 THEN
    FC_DL_ChuteFullPredict := -1.0; RETURN;   // 哨兵 -1：非有限或量纲越界 / Sentinel -1
END_IF
// 填充率域闸：0~100% 之外钳位
IF fFillPct < 0.0 THEN
    fFillPct := 0.0;                // 下限钳位 [%] / Clamp lower bound
ELSIF fFillPct > 100.0 THEN
    fFillPct := 100.0;              // 上限钳位 [%] / Clamp upper bound
END_IF
// 净流入：入流减出流，同量纲相减得 件/min（负值表示正在清空）
fNetPpm := fInflowPpm - fOutflowPpm;   // 净累积率 [件/min] / Net accumulation rate
// 剩余容量：容量 × (100 - 填充率) ÷ 100 = 件（% 约去，量纲自洽）
fRoomPcs := fCapacityPcs * ((100.0 - fFillPct) / 100.0); // 剩余容量 [件] / Remaining capacity [pcs]
// 净流正负双分支：净流非正时不溢出，给 0 与无风险标志
IF fNetPpm > 1.0E-9 THEN           // 净流分母显式零闸（R4/R21）/ Explicit zero gate on net rate
    // 件 ÷ (件/min) = min，×60 = s（量纲自洽）
    fTimeToFullS := fRoomPcs / fNetPpm * 60.0;  // 到满时间 [s] / Time to full [s]
    IF fTimeToFullS < 60.0 THEN
        xCritical := TRUE;          // 60 s 内将满料 / Will be full within 60 s
    END_IF
ELSE
    fTimeToFullS := 0.0;            // 净流非正，不会满料 / Net drain, never full
    xCritical    := FALSE;          // 无满料风险 / No full risk
END_IF
xValid := TRUE; FC_DL_ChuteFullPredict := fTimeToFullS;  // 返回到满时间 [s] / Return time to full
END_FUNCTION

(* ---- FC_DL_ClampDintChk.st ---- *)
(*==============================================================================
 * 名称 : FC_DL_ClampDintChk —— DINT 限幅 + 越界方向标志（nLo>nHi 判参数非法）
 * 分类 / 前缀 / 版本 : DL_Algo / FC_DL_ / 1.0.0
 * 溯源 : 开源语义参考（OSCAT/AixOCAT 族，MIT）或 clean-room IEC 实现，未复制源码
 * 平台 : 纯 IEC 61131-3
 * 功能说明 : 将 nIn 限幅到 [nLo,nHi] 并输出越界方向：nDir=-1 下限截断 /
 *            0 未截断 / +1 上限截断，供下游统计截断频次或触发量程告警。
 *            边界处理：nLo>nHi 判参数非法（区间为空），返回 0、nDir=0、
 *            bValid=FALSE 并置 eErr；nIn 恰等于边界值属未截断（nDir=0）。
 * 错误码 : 16#0001_1C05 = 区间非法（nLo>nHi，无合法限幅区间）
 *          eErr=0 且 bValid=TRUE 表示限幅结果与方向标志可用
 * 状态机 : R6 标注 N/A（纯函数无顺序状态，以本节替代 ELSE 兜底）
 * 红线 : R1/R2/R3 ✓ 零全局/零IO/纯IEC ｜ R4 ✓ 区间校验 ｜ R10 ✓ 标准转换 ｜ R11 ✓ 分号收尾 ｜ R15 ✓ 无保留字撞名
 * 修订记录 : 2026-11-23 v1.0.0 首次入库（R76）
 *============================================================================*)
FUNCTION FC_DL_ClampDintChk : DINT
VAR_INPUT
    nIn : DINT;    // 被限幅输入量 [-2147483648..2147483647] / input value to clamp
    nLo : DINT;    // 限幅下界（须 <=nHi）/ clamp lower bound, must be <= nHi
    nHi : DINT;    // 限幅上界（须 >=nLo）/ clamp upper bound, must be >= nLo
END_VAR
VAR_OUTPUT
    nDir   : INT;      // 越界方向 -1 下截断 / 0 未截断 / +1 上截断 / clamp direction
    eErr   : UDINT;    // 故障码，0=正常，1C05=区间非法 / error code, 0=ok, 1C05=invalid range
    bError : BOOL;     // TRUE=本件发生故障 / TRUE when fault occurred
    bValid : BOOL;     // TRUE=限幅结果可用 / TRUE when result is usable
END_VAR

FC_DL_ClampDintChk := 0;                     // 返回值预设 0 / preset return to zero
nDir   := 0;                                // 方向预设未截断 / preset direction to none
eErr   := 16#0000_0000;                     // 故障码清零 / clear error code
bError := FALSE;                            // 故障标志清零 / clear error flag
bValid := TRUE;                             // 预设输出可用 / preset valid flag

IF nLo > nHi THEN                           // 区间为空：参数非法 / empty range invalid
    eErr   := 16#0001_1C05;                 // 置区间非法码 / set invalid-range code
    bError := TRUE;                         // 置故障标志 / set error flag
    bValid := FALSE;                        // 输出不可用 / outputs not usable
    nDir   := 0;                            // 方向保持 0 / keep direction zero
    RETURN;                                 // 返回 0 / return zero
END_IF

IF nIn < nLo THEN                           // 低于下界 / below lower bound
    FC_DL_ClampDintChk := nLo;              // 截到下界 / clamp to lower bound
    nDir := -1;                             // 标记下限截断 / flag lower clamp
ELSIF nIn > nHi THEN                        // 高于上界 / above upper bound
    FC_DL_ClampDintChk := nHi;              // 截到上界 / clamp to upper bound
    nDir := 1;                              // 标记上限截断 / flag upper clamp
ELSE                                        // 区间内 / inside range
    FC_DL_ClampDintChk := nIn;              // 原值透传 / pass through
    nDir := 0;                              // 未截断 / not clamped
END_IF

END_FUNCTION

(* ---- FC_DL_CoilDiameterCalc.st ---- *)
(*==============================================================================
 * 组件名称 (Component)  : FC_DL_CoilDiameterCalc
 * 所属子库 (Sublibrary) : DL_Algo
 * 当前版本 (Version)    : 1.0.0
 * 组件分类 (Category)   : 函数（FUNCTION）· 纯函数 · 卷绕工艺量反算
 * 兼容性   (Platform)   : CODESYS 3.5 / TwinCAT 3 / 汇川 InoProShop / Schneider
 *                         Machine Expert；仅用标准算术、ABS、LIMIT
 * 功能描述 (Function)   : 由「材料线速度 + 卷轴转速 + 机械传动比」反算瞬时卷径
 *                         直径 = 线速度 乘以 传动比 除以 (派 乘以 转速)，并同时
 *                         给出卷径变化率与相对卷芯的累计层数。是收放卷张力控制
 *                         （扭矩等于张力乘卷径除二）、线速度匹配、排线节距计算
 *                         的数据源头。
 * 与既有件边界 (Boundary): 本件只做瞬时几何反算（无状态、无记忆）；层厚积分
 *                         递推与排线执行属 FB_DL_WindingTraverse 的职责；两者
 *                         互为校验关系（可把本件结果注入该块的注入卷径引脚做
 *                         比对），但代码零调用、零耦合，禁止在本件内调用任何
 *                         功能块。
 * 设计要点 (Key notes)  : ① 低速保护是核心工程语义：转速低于 0.5 转每分时
 *                           编码器低频量化会让反算卷径跳动到毫米级，此时沿用
 *                           上次有效卷径而不是归零。停机瞬间卷径突然归零会让
 *                           张力给定瞬间飙到上限，是现场最常见的事故源；
 *                         ② 卷芯保护：反算卷径小于卷芯直径说明打滑或测速错，
 *                           按卷芯直径修正并置码，绝不把几何上不可能的值下发；
 *                         ③ 一阶低通首拍无滞后：上次卷径为 0 时直接取原始值，
 *                           避免从 0 缓慢爬升（R19 精神）；
 *                         ④ 变化率先算再更新历史值，次序颠倒会得到恒 0；
 *                         ⑤ 所有除法分母（转速、滤波时间常数加周期、上次卷径、
 *                           厚度）均有守卫或常量域保证，无除零面。
 * 开源溯源 (Origin)     : lgf-technology。参考 LGF（Libre Graphical Framework）
 *                         公开函数库「Technology」分类中卷绕类函数的功能分类
 *                         与参数域（线速度 / 转速 / 传动比 三段入口形态），只借
 *                         分类、参数域与命名习惯，公式重排与实现 100% 自有
 *                         clean-room，不构成衍生作品。
 * 依赖     (Depends)    : 无 DL_ 内部依赖；无标准库功能块依赖
 * 故障码表 (Error codes):
 *   16#0002_1D01【信息级】线速度越界被钳位
 *   16#0002_1D02【信息级】传动比越界被钳位
 *   16#0002_1D03【信息级】卷芯直径或材料厚度越界被钳位
 *   16#0002_1D04【信息级】反算卷径小于卷芯直径，已按卷芯修正（疑似打滑）
 *   16#0002_1D10【信息级】转速过低不可信或入参非有限，沿用上次有效值
 * 验收向量 (Acceptance) :
 *   V1 线速度 100 米每分 / 转速 100 转每分 / 传动比 1 → 卷径约 0.3183 米
 *   V2 转速 0.2 转每分（低于 0.5）→ 返回上次卷径、变化率 0、码 1D10
 *   V3 线速度 10 / 转速 100 / 卷芯 0.2 → 原始值 0.0318 小于卷芯，修正为 0.2
 *      并置 1D04
 *   V4 上次卷径 0 且滤波使能 → 首拍输出等于原始值（无滞后）
 *   V5 上次卷径 0.3 / 当前 0.302 / 周期 0.01 → 变化率 0.2 米每秒
 * 红线自检 (Redline)    : R1 零全局变量表与外部变量引用 ｜ R2 零物理地址直写
 *                         R3 纯 IEC 61131-3 ｜ R4 全部除法分母有守卫、浮点判等
 *                         用容差、非有限值筛查 ｜ R5 全变量中英双语同行注释
 *                         R6 N/A（纯函数）｜ R7 N/A（无实例调用）
 * 修订历史 (Revision)   :
 *   2026-11-15  v1.0.0  首版入库（Round 10 · 工艺物理量链）
 *============================================================================*)

FUNCTION FC_DL_CoilDiameterCalc : LREAL
VAR_INPUT
    fLineSpeed : LREAL := 0.0;      // 材料线速度，域 0 到 3000 [米每分] / Material line speed, 0 to 3000 metres per minute
    fShaftRpm  : LREAL := 0.0;      // 卷轴转速，域 0 到 6000，低于 0.5 视为停机 [转每分] / Shaft speed, below 0.5 rpm treated as standstill
    fGearRatio : LREAL := 1.0;      // 卷轴对电机传动比，域 0.01 到 1000，1.0 为直连 [-] / Shaft to motor gear ratio, 1.0 means direct drive
    fCoreDia   : LREAL := 0.100;    // 卷芯（纸管）直径，域 0.01 到 1.0 [米] / Core diameter, 0.01 to 1.0 m
    fThickness : LREAL := 0.0001;   // 材料厚度，域 1 微米到 10 毫米，层数积分用 [米] / Material thickness, used by the layer count
    fPrevDia   : LREAL := 0.0;      // 上拍卷径，0 表示无历史（变化率出口置 0）[米] / Previous diameter, 0 means no history
    fTaskCycle : LREAL := 0.01;     // 任务周期，域 1 毫秒到 1 秒，变化率换算用 [s] / Task cycle time
    bFilterEn  : BOOL := TRUE;      // 一阶低通使能，用于抑制编码器量化噪声 [-] / First-order low-pass enable
    fFilterTau : LREAL := 1.0;      // 低通时间常数，域 0.1 到 10 [s] / Low-pass time constant
END_VAR
VAR_OUTPUT
    fDia        : LREAL;    // 估算卷径，低通使能时为滤波后的值 [米] / Estimated diameter, filtered when enabled
    fDiaRaw     : LREAL;    // 未滤波原始卷径，用于诊断与比对 [米] / Unfiltered diameter for diagnostics
    fDiaRate    : LREAL;    // 卷径变化率，正值为收卷增大 [米每秒] / Diameter rate, positive when winding up
    fLayerCount : LREAL;    // 相对卷芯的累计层数，由厚度推算 [层] / Layer count relative to the core
    bValid      : BOOL;     // 计算有效，任一钳位或修正事件为 FALSE [-] / TRUE when no clamping or correction happened
    uErrorId    : UDINT;    // 事件码，0 = 无事件 / Event code, 0 = no event
END_VAR
VAR
    fGearUse  : LREAL;      // 生效传动比（已钳位）[-] / Effective gear ratio
    fCoreUse  : LREAL;      // 生效卷芯直径（已钳位）[米] / Effective core diameter
    fThickUse : LREAL;      // 生效材料厚度（已钳位）[米] / Effective thickness
    fLineUse  : LREAL;      // 生效线速度（已钳位）[米每分] / Effective line speed
    fDtUse    : LREAL;      // 生效任务周期（已钳位）[s] / Effective task cycle
    fTauUse   : LREAL;      // 生效滤波时间常数（已钳位）[s] / Effective filter time constant
    fAlpha    : LREAL;      // 一阶低通权重 [-] / First-order filter weight
    bDirty    : BOOL;       // 是否发生过钳位或修正事件 [-] / TRUE when any clamp or correction fired
END_VAR
VAR CONSTANT
    DL_PI         : LREAL := 3.141592653589793;  // 圆周率 [-] / Pi
    DL_SEC_PER_MIN: LREAL := 60.0;               // 分钟转秒 [s每分] / Seconds per minute
    DL_VMAX       : LREAL := 3000.0;             // 线速度上限，约 50 米每秒，覆盖高速分切 [米每分] / Line speed upper bound
    DL_NMAX       : LREAL := 6000.0;             // 转速上限 [转每分] / Shaft speed upper bound
    DL_RPM_EPS    : LREAL := 0.5;                // 转速判零门限，低于此不反算 [转每分] / Speed floor below which the inverse is untrustworthy
    DL_DIA_MIN    : LREAL := 0.01;               // 卷径下限 [米] / Diameter lower bound
    DL_DIA_MAX    : LREAL := 3.0;                // 卷径上限 [米] / Diameter upper bound
    DL_CORE_MIN   : LREAL := 0.01;               // 卷芯直径下限 [米] / Core diameter lower bound
    DL_CORE_MAX   : LREAL := 1.0;                // 卷芯直径上限 [米] / Core diameter upper bound
    DL_THICK_MIN  : LREAL := 1.0E-6;             // 厚度下限，1 微米 [米] / Thickness lower bound
    DL_THICK_MAX  : LREAL := 0.01;               // 厚度上限，10 毫米 [米] / Thickness upper bound
    DL_GEAR_MIN   : LREAL := 0.01;               // 传动比下限 [-] / Gear ratio lower bound
    DL_GEAR_MAX   : LREAL := 1000.0;             // 传动比上限 [-] / Gear ratio upper bound
    DL_TAU_MIN    : LREAL := 0.1;                // 滤波时间常数下限 [s] / Filter time constant lower bound
    DL_TAU_MAX    : LREAL := 10.0;               // 滤波时间常数上限 [s] / Filter time constant upper bound
    DL_CYCLE_MIN  : LREAL := 0.001;              // 任务周期下限 [s] / Task cycle lower bound
    DL_CYCLE_MAX  : LREAL := 1.0;                // 任务周期上限 [s] / Task cycle upper bound
    DL_FLOAT_EPS  : LREAL := 1.0E-9;             // 浮点容差 [-] / Float tolerance
    DL_BIG        : LREAL := 1.0E300;            // 非有限值兜底门限 [-] / Magnitude guard
    DL_LAYER_DIV  : LREAL := 2.0;                // 层数公式中的二倍因子，单层增径为两倍厚度 [-] / Two-times factor of the layer formula
END_VAR

(*------------------------------------------------------------------------------
 * 段 1｜输出预置
 *      Pre-set outputs
 *-----------------------------------------------------------------------------*)
FC_DL_CoilDiameterCalc := 0.0;
fDia        := 0.0;
fDiaRaw     := 0.0;
fDiaRate    := 0.0;
fLayerCount := 0.0;
bValid      := FALSE;
uErrorId    := 16#0000_0000;
bDirty      := FALSE;

(*------------------------------------------------------------------------------
 * 段 2｜入参有限性筛查（边界 B1）：任一非有限即按不可信处理，沿用上次值
 *      Input finiteness check: any non-finite value is untrusted
 *-----------------------------------------------------------------------------*)
IF (fLineSpeed <> fLineSpeed) OR (fShaftRpm <> fShaftRpm) OR (fGearRatio <> fGearRatio)
   OR (fCoreDia <> fCoreDia) OR (fThickness <> fThickness) OR (fPrevDia <> fPrevDia)
   OR (fTaskCycle <> fTaskCycle) OR (fFilterTau <> fFilterTau) THEN
    fDia     := fPrevDia;            // 沿用上次有效卷径，绝不归零
    fDiaRaw  := fPrevDia;
    fDiaRate := 0.0;
    uErrorId := 16#0002_1D10;
    RETURN;
END_IF

IF (ABS(fLineSpeed) > DL_BIG) OR (ABS(fShaftRpm) > DL_BIG) OR (ABS(fPrevDia) > DL_BIG) THEN
    fDia     := fPrevDia;
    fDiaRaw  := fPrevDia;
    fDiaRate := 0.0;
    uErrorId := 16#0002_1D10;
    RETURN;
END_IF

(*------------------------------------------------------------------------------
 * 段 3｜参数域钳位（信息级）：钳位后继续计算，宁可给近似值也不给 0 断链
 *      Parameter clamping with informational codes, computation always continues
 *-----------------------------------------------------------------------------*)
fLineUse := fLineSpeed;
IF fLineUse < 0.0 THEN
    fLineUse := 0.0;
    uErrorId := 16#0002_1D01;
    bDirty   := TRUE;
ELSIF fLineUse > DL_VMAX THEN
    fLineUse := DL_VMAX;
    uErrorId := 16#0002_1D01;
    bDirty   := TRUE;
END_IF

fGearUse := fGearRatio;
IF fGearUse < DL_GEAR_MIN THEN
    fGearUse := DL_GEAR_MIN;
    uErrorId := 16#0002_1D02;
    bDirty   := TRUE;
ELSIF fGearUse > DL_GEAR_MAX THEN
    fGearUse := DL_GEAR_MAX;
    uErrorId := 16#0002_1D02;
    bDirty   := TRUE;
END_IF

fCoreUse := fCoreDia;
IF fCoreUse < DL_CORE_MIN THEN
    fCoreUse := DL_CORE_MIN;
    uErrorId := 16#0002_1D03;
    bDirty   := TRUE;
ELSIF fCoreUse > DL_CORE_MAX THEN
    fCoreUse := DL_CORE_MAX;
    uErrorId := 16#0002_1D03;
    bDirty   := TRUE;
END_IF

fThickUse := fThickness;
IF fThickUse < DL_THICK_MIN THEN
    fThickUse := DL_THICK_MIN;
    uErrorId  := 16#0002_1D03;
    bDirty    := TRUE;
ELSIF fThickUse > DL_THICK_MAX THEN
    fThickUse := DL_THICK_MAX;
    uErrorId  := 16#0002_1D03;
    bDirty    := TRUE;
END_IF

fDtUse := fTaskCycle;
IF fDtUse < DL_CYCLE_MIN THEN
    fDtUse := DL_CYCLE_MIN;
ELSIF fDtUse > DL_CYCLE_MAX THEN
    fDtUse := DL_CYCLE_MAX;
END_IF

fTauUse := fFilterTau;
IF fTauUse < DL_TAU_MIN THEN
    fTauUse := DL_TAU_MIN;
ELSIF fTauUse > DL_TAU_MAX THEN
    fTauUse := DL_TAU_MAX;
END_IF

(*------------------------------------------------------------------------------
 * 段 4｜低速保护（关键工程语义，边界 B2）：转速低于门限不反算，沿用上次值
 *      Low-speed protection: below the speed floor the inverse is skipped
 *      现场理由：停机瞬间反算卷径会突然塌到接近 0，若直接下发会让张力扭矩
 *      给定瞬间飙到上限，是收放卷最常见的断料与飞车诱因
 *-----------------------------------------------------------------------------*)
IF fShaftRpm < DL_RPM_EPS THEN
    fDia     := fPrevDia;                          // 沿用上次有效卷径
    fDiaRaw  := fPrevDia;
    fDiaRate := 0.0;
    uErrorId := 16#0002_1D10;
    IF fPrevDia >= DL_DIA_MIN THEN
        bValid := TRUE;                            // 有历史值时结果仍可用
    ELSE
        bValid := FALSE;                           // 无历史值时结果不可用
    END_IF
    FC_DL_CoilDiameterCalc := fDia;
    RETURN;
END_IF

(*------------------------------------------------------------------------------
 * 段 5｜主反算：直径 = 线速度 乘以 传动比 除以 (派 乘以 转速)
 *      Main inverse: diameter equals line speed times ratio over pi times rpm
 *      写法一（保留单位可读性，分子分母同除 60）：
 *        原始值 = (线速度 除以 60) 乘以 传动比 除以 (派 乘以 (转速 除以 60))
 *      化简后等价于：原始值 = 线速度 乘以 传动比 除以 (派 乘以 转速)
 *      两式完全等价，此处按写法一书写以便维护者核对量纲，禁止改成其它形式
 *      分母的转速已由段 4 保证不小于 0.5，派为常量，无除零面
 *-----------------------------------------------------------------------------*)
fDiaRaw := (fLineUse / DL_SEC_PER_MIN) * fGearUse
           / (DL_PI * (fShaftRpm / DL_SEC_PER_MIN));

(*------------------------------------------------------------------------------
 * 段 6｜卷芯保护与卷径钳位（边界 B3）：几何上不可能的值必须修正
 *      Core protection and diameter clamping: geometrically impossible values fixed
 *-----------------------------------------------------------------------------*)
IF fDiaRaw < fCoreUse THEN
    fDiaRaw  := fCoreUse;          // 卷径不可能小于卷芯：疑似打滑或测速错
    uErrorId := 16#0002_1D04;
    bDirty   := TRUE;
END_IF

fDiaRaw := LIMIT(DL_DIA_MIN, fDiaRaw, DL_DIA_MAX);

(*------------------------------------------------------------------------------
 * 段 7｜一阶低通（首拍无滞后）：分母恒大于 0.1，无除零面
 *      First-order low pass with no lag on the first cycle
 *-----------------------------------------------------------------------------*)
IF bFilterEn THEN
    IF fPrevDia < DL_FLOAT_EPS THEN
        fDia := fDiaRaw;                            // 首拍直接取原始值，避免从 0 爬升
    ELSE
        fAlpha := fDtUse / (fTauUse + fDtUse);      // 分母不小于 0.101
        fDia   := fPrevDia + fAlpha * (fDiaRaw - fPrevDia);
    END_IF
ELSE
    fDia := fDiaRaw;
END_IF

fDia := LIMIT(DL_DIA_MIN, fDia, DL_DIA_MAX);

(*------------------------------------------------------------------------------
 * 段 8｜变化率（先算再更新历史值，次序写死）
 *      Diameter rate computed before the history value is refreshed
 *-----------------------------------------------------------------------------*)
IF fPrevDia > DL_FLOAT_EPS THEN
    fDiaRate := (fDia - fPrevDia) / fDtUse;         // 周期已被钳到不小于 1 毫秒
ELSE
    fDiaRate := 0.0;                                // 无历史值时不产生变化率
END_IF

(*------------------------------------------------------------------------------
 * 段 9｜层数：单层增径为两倍厚度，故层数等于半径差除以厚度
 *      Layer count: each layer adds two thicknesses to the diameter
 *-----------------------------------------------------------------------------*)
fLayerCount := (fDia - fCoreUse) / (DL_LAYER_DIV * fThickUse);

IF fLayerCount < 0.0 THEN
    fLayerCount := 0.0;                             // 层数不得为负（卷芯修正后的边界）
END_IF

(*------------------------------------------------------------------------------
 * 段 10｜有效性与返回值收口
 *      Validity and return value close-out
 *-----------------------------------------------------------------------------*)
IF bDirty THEN
    bValid := FALSE;                                // 发生过钳位或修正，结果标注为近似
ELSE
    bValid := TRUE;
END_IF

FC_DL_CoilDiameterCalc := fDia;
END_FUNCTION

(* ---- FC_DL_ContainerStackHeightCalc.st ---- *)
(*
 * FC_DL_ContainerStackHeightCalc | C2 | DL_Algo
 * 功能：堆场贝位层高与箱位换算（顶面标高、剩余层数、超高判定）       单位：层 [1]、层高 [m]、标高 [m]
 * 工况边界：nTier 须落在 [1, nMaxTier] 且 nMaxTier≥1，否则判故障 9611 并输出安全值（超高置 TRUE 阻止堆箱）；堆高上限 rMaxStackHm 须 >0；层高须 >0 且有限
 * 代数值回代：nTier=5、rTierHm=2.591、rBaseHm=0.30 → top=0.30+4×2.591+2.591=13.255 m（spec 记 13.25 m，取两位小数一致）
 * 开源溯源：clean-room 自研，未复制任何第三方代码（无外部来源）
 *)
FUNCTION FC_DL_ContainerStackHeightCalc : BOOL
VAR_INPUT
    nTier        : INT;              // 目标层号（1 起）| target tier, one based [层]
    nMaxTier     : INT;              // 该贝位允许的最大层数 | maximum tier count of this bay [层]
    rTierHm      : REAL := 2.591;    // 单层箱高（含层间间隙）| container height including the gap [m]
    rBaseHm      : REAL := 0.30;     // 基础标高（码头面至第一层箱底）| base elevation from the quay to the first box bottom [m]
    rMaxStackHm  : REAL := 30.0;     // 堆场允许最大标高 | maximum permitted stack elevation [m]
END_VAR
VAR_OUTPUT
    rTopElevM  : REAL;               // 目标层顶面标高 | top elevation of the target tier [m]
    nFreeTier  : INT;                // 剩余可用层数 | remaining tier capacity [层]
    xOverHeight: BOOL;               // 超高（顶面超 rMaxStackHm）| over height, the top exceeds rMaxStackHm
    xValid     : BOOL;               // 输出有效 | outputs valid
    nFaultCode : INT;                // 0=无 / 9611=层号或配置非法 | 0 none, 9611 illegal tier or configuration
END_VAR
VAR
    xFinTierH : BOOL;                // 层高有限性 | tier height is finite
    xFinBase  : BOOL;                // 基础标高有限性 | base elevation is finite
    xFinMaxH  : BOOL;                // 堆高上限有限性 | stack height limit is finite
END_VAR
VAR CONSTANT
    DL_CSH_TOL_M : REAL := 1.0E-6;   // 浮点比较容差 | floating comparison tolerance [m]
END_VAR

// 段1｜非有限闸（R19）
xFinTierH := (rTierHm = rTierHm) AND ((rTierHm - rTierHm) = 0.0);
xFinBase := (rBaseHm = rBaseHm) AND ((rBaseHm - rBaseHm) = 0.0);
xFinMaxH := (rMaxStackHm = rMaxStackHm) AND ((rMaxStackHm - rMaxStackHm) = 0.0);
IF (NOT xFinTierH) OR (NOT xFinBase) OR (NOT xFinMaxH) THEN
    rTopElevM := 0.0;                // 安全值：标高 0 | safe value, zero elevation
    nFreeTier := 0;                  // 安全值：无剩余层 | safe value, no capacity left
    xOverHeight := TRUE;             // 安全值：判超高，禁止堆箱 | safe value, over height so stacking is blocked
    xValid := FALSE;
    nFaultCode := 9611;
    FC_DL_ContainerStackHeightCalc := FALSE;
    RETURN;
END_IF

// 段2｜域闸：层号范围与几何配置（先判后用）
IF (nMaxTier < 1) OR (nTier < 1) OR (nTier > nMaxTier)
   OR (rTierHm <= 0.0) OR (rMaxStackHm <= 0.0) THEN
    rTopElevM := 0.0;
    nFreeTier := 0;
    xOverHeight := TRUE;
    xValid := FALSE;
    nFaultCode := 9611;
    FC_DL_ContainerStackHeightCalc := FALSE;
    RETURN;
END_IF

// 段3｜算法：top = base + (tier-1)*tierH + tierH
rTopElevM := rBaseHm + INT_TO_REAL(nTier - 1) * rTierHm + rTierHm;
nFreeTier := nMaxTier - nTier;                          // 剩余层数（同型整数运算，无跨型转换）| remaining tiers, same integer type
IF nFreeTier < 0 THEN
    nFreeTier := 0;                                     // 保险钳位（段2已保证非负）| defensive clamp
END_IF

// 段4｜超高判定：用未截断的原始标高与限值直接比较
xOverHeight := rTopElevM > (rMaxStackHm + DL_CSH_TOL_M);
nFaultCode := 0;
xValid := TRUE;
FC_DL_ContainerStackHeightCalc := TRUE;
END_FUNCTION

(* ---- FC_DL_CraneCycleTimeEstimate.st ---- *)
(*
 * FC_DL_CraneCycleTimeEstimate | C2 | DL_Algo
 * 功能：单箱作业循环时间估算（起升 / 小车 / 大车三轴 + 固定辅助时间）       单位：距离 [m]、速度 [m/s]、加速度 [m/s²]、时间 [s]
 * 工况边界：各轴速度与加速度须 >0 且有限；某轴距离 ≤0 视为该轴不动作，时间计 0；含加速与减速的对称梯形近似，不含防摇等待与人工对箱时间（由 rFixedS 覆盖）
 * 代数值回代：起升 20 m/1.2+1.2/0.5=19.07 s；小车 30/2.5+2.5/0.5=17.0 s；大车 0 s；总=19.07+17.0+0+25=61.07 s（spec 记 19.1/17.0/0/61.1 s，一致）
 * 开源溯源：clean-room 自研，未复制任何第三方代码（无外部来源）
 *)
FUNCTION FC_DL_CraneCycleTimeEstimate : BOOL
VAR_INPUT
    rHoistDistM   : REAL := 20.0;    // 起升行程 | hoist travel [m]
    rTrolleyDistM : REAL := 30.0;    // 小车行程 | trolley travel [m]
    rGantryDistM  : REAL := 0.0;     // 大车行程（单箱作业常为 0）| gantry travel, usually zero per box [m]
    rVHoist       : REAL := 1.2;     // 起升额定速度 | hoist rated speed [m/s]
    rVTrolley     : REAL := 2.5;     // 小车额定速度 | trolley rated speed [m/s]
    rVGantry      : REAL := 3.0;     // 大车额定速度 | gantry rated speed [m/s]
    rAcc          : REAL := 0.5;     // 统一加减速度 | common acceleration and deceleration [m/s²]
    rFixedS       : REAL := 25.0;    // 固定辅助时间（对箱、开闭锁等）| fixed handling time [s]
END_VAR
VAR_OUTPUT
    rHoistS   : REAL;                // 起升轴时间 | hoist axis time [s]
    rTrolleyS : REAL;                // 小车轴时间 | trolley axis time [s]
    rGantryS  : REAL;                // 大车轴时间 | gantry axis time [s]
    rCycleS   : REAL;                // 循环总时间 | total cycle time [s]
    xValid    : BOOL;                // 输出有效 | outputs valid
END_VAR
VAR
    xFinH     : BOOL;                // 起升行程有限性 | hoist travel is finite
    xFinT     : BOOL;                // 小行程有限性 | trolley travel is finite
    xFinG     : BOOL;                // 大车行程有限性 | gantry travel is finite
    xFinVh    : BOOL;                // 起升速度有限性 | hoist speed is finite
    xFinVt    : BOOL;                // 小车速度有限性 | trolley speed is finite
    xFinVg    : BOOL;                // 大车速度有限性 | gantry speed is finite
    xFinA     : BOOL;                // 加速度有限性 | acceleration is finite
    xFinFixed : BOOL;                // 固定时间有限性 | fixed time is finite
    rCritH    : REAL;                // 起升达到额定速度所需行程 | travel needed to reach the hoist rated speed [m]
    rCritT    : REAL;                // 小车达到额定速度所需行程 | travel needed to reach the trolley rated speed [m]
    rCritG    : REAL;                // 大车达到额定速度所需行程 | travel needed to reach the gantry rated speed [m]
END_VAR

// 段1｜非有限闸（R19）
xFinH := (rHoistDistM = rHoistDistM) AND ((rHoistDistM - rHoistDistM) = 0.0);
xFinT := (rTrolleyDistM = rTrolleyDistM) AND ((rTrolleyDistM - rTrolleyDistM) = 0.0);
xFinG := (rGantryDistM = rGantryDistM) AND ((rGantryDistM - rGantryDistM) = 0.0);
xFinVh := (rVHoist = rVHoist) AND ((rVHoist - rVHoist) = 0.0);
xFinVt := (rVTrolley = rVTrolley) AND ((rVTrolley - rVTrolley) = 0.0);
xFinVg := (rVGantry = rVGantry) AND ((rVGantry - rVGantry) = 0.0);
xFinA := (rAcc = rAcc) AND ((rAcc - rAcc) = 0.0);
xFinFixed := (rFixedS = rFixedS) AND ((rFixedS - rFixedS) = 0.0);
IF (NOT xFinH) OR (NOT xFinT) OR (NOT xFinG) OR (NOT xFinVh) OR (NOT xFinVt)
   OR (NOT xFinVg) OR (NOT xFinA) OR (NOT xFinFixed) THEN
    rHoistS := 0.0;                  // 安全值：时间全 0 | safe value, all zero
    rTrolleyS := 0.0;
    rGantryS := 0.0;
    rCycleS := 0.0;
    xValid := FALSE;
    FC_DL_CraneCycleTimeEstimate := FALSE;
    RETURN;
END_IF

// 段2｜域闸：速度与加速度必须为正（速度在分母）；固定时间不得为负
IF (rVHoist <= 0.0) OR (rVTrolley <= 0.0) OR (rVGantry <= 0.0)
   OR (rAcc <= 0.0) OR (rFixedS < 0.0) THEN
    rHoistS := 0.0;
    rTrolleyS := 0.0;
    rGantryS := 0.0;
    rCycleS := 0.0;
    xValid := FALSE;
    FC_DL_CraneCycleTimeEstimate := FALSE;
    RETURN;
END_IF

// 段3｜起升轴：d ≥ v²/a 走梯形 t=d/v+v/a，否则三角形 t=2·SQRT(d/a)
rCritH := (rVHoist * rVHoist) / rAcc;
IF rHoistDistM <= 0.0 THEN
    rHoistS := 0.0;                                          // 该轴不动作 | axis not moving
ELSIF rHoistDistM >= rCritH THEN
    rHoistS := rHoistDistM / rVHoist + rVHoist / rAcc;
ELSE
    rHoistS := 2.0 * SQRT(rHoistDistM / rAcc);
END_IF

// 段4｜小车轴
rCritT := (rVTrolley * rVTrolley) / rAcc;
IF rTrolleyDistM <= 0.0 THEN
    rTrolleyS := 0.0;
ELSIF rTrolleyDistM >= rCritT THEN
    rTrolleyS := rTrolleyDistM / rVTrolley + rVTrolley / rAcc;
ELSE
    rTrolleyS := 2.0 * SQRT(rTrolleyDistM / rAcc);
END_IF

// 段5｜大车轴
rCritG := (rVGantry * rVGantry) / rAcc;
IF rGantryDistM <= 0.0 THEN
    rGantryS := 0.0;
ELSIF rGantryDistM >= rCritG THEN
    rGantryS := rGantryDistM / rVGantry + rVGantry / rAcc;
ELSE
    rGantryS := 2.0 * SQRT(rGantryDistM / rAcc);
END_IF

// 段6｜总时间与出口
rCycleS := rHoistS + rTrolleyS + rGantryS + rFixedS;
xValid := TRUE;
FC_DL_CraneCycleTimeEstimate := TRUE;
END_FUNCTION

(* ---- FC_DL_CraneLoadMomentCalc.st ---- *)
(*
 * FC_DL_CraneLoadMomentCalc | C2 | DL_Algo
 * 功能：载荷倾覆力矩、抗倾覆力矩与安全系数（含重心偏移附加判据）       单位：质量 [t]、长度 [m]、力矩 [t·m]、安全系数 [1]
 * 工况边界：抗倾覆力矩采用 spec 简化式 Mr=W_crane×轮距/2（整机按最不利支腿回转取轮距半宽）；重心偏移 rCgDistM 仅作为附加稳定判据（超过轮距半宽即判不安全），不进入 Mr 计算；吊重与跨距须 >0 且有限
 * 代数值回代：load=40 t @40 m → Mo=1600 t·m；crane=1000 t、轮距 16 m → Mr=1000×8=8000 t·m；SF=8000/1600=5.0 ≥1.5 → xSafe=TRUE（与 spec 回代行一致）
 * 开源溯源：clean-room 自研，未复制任何第三方代码（无外部来源）
 *)
FUNCTION FC_DL_CraneLoadMomentCalc : BOOL
VAR_INPUT
    rLoadT        : REAL;            // 吊重（含吊具）| lifted load including the spreader [t]
    rOutreachM    : REAL;            // 工作幅度（回转中心至吊重）| working outreach [m]
    rCraneWeightT : REAL;            // 整机自重 | crane dead weight [t]
    rCgDistM      : REAL;            // 整机重心至回转中心距离 | centre of gravity offset from the slew centre [m]
    rWheelBaseM   : REAL := 16.0;    // 大车轮距（轨距）| rail gauge or wheel base [m]
    rSfMin        : REAL := 1.5;     // 要求最小抗倾覆安全系数 | required minimum safety factor [1]
END_VAR
VAR_OUTPUT
    rOverturnMomentTm : REAL;        // 倾覆力矩 Mo | overturning moment [t·m]
    rResistMomentTm   : REAL;        // 抗倾覆力矩 Mr | resisting moment [t·m]
    rSafetyFactor     : REAL;        // 安全系数 SF=Mr/Mo | safety factor [1]
    xSafe             : BOOL;        // 稳定判定（SF≥限值 且 重心不越界）| stable verdict
    xCgOverLimit      : BOOL;        // 重心偏移越界（信息级）| centre of gravity out of range, informational
    xValid            : BOOL;        // 输出有效 | outputs valid
END_VAR
VAR
    xFinLoad  : BOOL;                // 吊重有限性 | load is finite
    xFinOut   : BOOL;                // 幅度有限性 | outreach is finite
    xFinW     : BOOL;                // 自重有限性 | dead weight is finite
    xFinCg    : BOOL;                // 重心偏移有限性 | centre of gravity offset is finite
    xFinWb    : BOOL;                // 轮距有限性 | wheel base is finite
    xFinSf    : BOOL;                // 安全系数限值有限性 | safety factor limit is finite
END_VAR
VAR CONSTANT
    DL_CLM_EPS : REAL := 1.0E-9;     // 除零保护阈值 | division guard threshold [t·m]
END_VAR

// 段1｜非有限闸（R19）
xFinLoad := (rLoadT = rLoadT) AND ((rLoadT - rLoadT) = 0.0);
xFinOut := (rOutreachM = rOutreachM) AND ((rOutreachM - rOutreachM) = 0.0);
xFinW := (rCraneWeightT = rCraneWeightT) AND ((rCraneWeightT - rCraneWeightT) = 0.0);
xFinCg := (rCgDistM = rCgDistM) AND ((rCgDistM - rCgDistM) = 0.0);
xFinWb := (rWheelBaseM = rWheelBaseM) AND ((rWheelBaseM - rWheelBaseM) = 0.0);
xFinSf := (rSfMin = rSfMin) AND ((rSfMin - rSfMin) = 0.0);
IF (NOT xFinLoad) OR (NOT xFinOut) OR (NOT xFinW) OR (NOT xFinCg)
   OR (NOT xFinWb) OR (NOT xFinSf) THEN
    rOverturnMomentTm := 0.0;        // 安全值：力矩 0 | safe value, zero moments
    rResistMomentTm := 0.0;
    rSafetyFactor := 0.0;            // 安全值：安全系数 0（判不稳）| safe value, zero factor means unstable
    xSafe := FALSE;
    xCgOverLimit := TRUE;
    xValid := FALSE;
    FC_DL_CraneLoadMomentCalc := FALSE;
    RETURN;
END_IF

// 段2｜域闸：吊重与幅度必须为正（Mo 入分母），轮距与安全系数限值必须为正
IF (rLoadT <= 0.0) OR (rOutreachM <= 0.0) OR (rWheelBaseM <= 0.0) OR (rSfMin <= 0.0) THEN
    rOverturnMomentTm := 0.0;
    rResistMomentTm := 0.0;
    rSafetyFactor := 0.0;
    xSafe := FALSE;
    xCgOverLimit := TRUE;
    xValid := FALSE;
    FC_DL_CraneLoadMomentCalc := FALSE;
    RETURN;
END_IF

// 段3｜力矩：Mo = W_load×L_out；Mr = W_crane×轮距/2（spec 简化式）
rOverturnMomentTm := rLoadT * rOutreachM;
rResistMomentTm := rCraneWeightT * (rWheelBaseM / 2.0);

// 段4｜安全系数：分母 Mo 已由段2保证 >0，仍按阈值显式防零
IF rOverturnMomentTm > DL_CLM_EPS THEN
    rSafetyFactor := rResistMomentTm / rOverturnMomentTm;
ELSE
    rSafetyFactor := 0.0;            // 理论上不可达（段2已排除），防御性兜底 | unreachable defence
END_IF

// 段5｜稳定判定：安全系数达标 且 重心不越轮距半宽（判据与出口同源于原始输入）
xCgOverLimit := rCgDistM > (rWheelBaseM / 2.0 + 1.0E-6);
xSafe := (rSafetyFactor >= rSfMin) AND (NOT xCgOverLimit);
xValid := TRUE;
FC_DL_CraneLoadMomentCalc := TRUE;
END_FUNCTION

(* ---- FC_DL_DeadtimeTapCalc.st ---- *)
//==============================================================================
// 函数：FC_DL_DeadtimeTapCalc ｜ 中文名称：死区时间→离散拍数向上取整换算
// 所属子库：DL_Algo ｜ 版本：v1.0.0 ｜ 日期：2026-11-23
// 兼容：CODESYS V3.5+ / TwinCAT 3 / 汇川 InoProShop（纯标准库）
// 功能描述：nTicks = CEIL(tDeadtime / tSample) 换算原子（Smith 预估器/
//           死区补偿前置）。取整纪律（终审必查项）：禁 TRUNC(x)+1 写法——
//           先 TRUNC 得整商，再按余量 > 容差进位；整商已达 DINT 上限且仍有
//           余量时饱和钳位 + bSaturated 声明（防进位溢出回绕）。
//           分工声明：离散拍数原子属本件；Smith 预估本体属
//           FB_DL_SmithPredictor，互不替代。
// 开源溯源 (Origin)：原创实现（自研-std 标准包装线，零外部源码行，clean-room
//           独立编写）
// 公开接口清单：输入 tDeadtime / tSample；输出 nTicks / bSaturated / bValid
// 错误码表：纯函数无状态机码轨；无效输入经 bValid = FALSE 表达（哨兵返回
//           0），饱和经 bSaturated 声明，本件不占用 16#0002 段码位
// 状态机：N/A（纯函数，无状态，可重入）
// 边界行为：① tSample <= 0（采样拍长非法）→ 拒绝（哨兵 0 返回）；
//           ② tDeadtime < 0 → 拒绝；tDeadtime = 0 合法（nTicks = 0）；
//           ③ 余量 > 1.0E-6 才进位（纯整除不虚进一位）；
//           ④ 商超 DINT 上限且有进位需求 → 饱和钳 2147483647 + bSaturated；
//           ⑤ 非有限输入 → 哨兵 0 返回。
// 修订历史：v1.0.0 2026-11-23 首版（R73 派单 · 批 3 · 序 18）
//==============================================================================

(*------------------------------------------------------------------------------
 * 调用示例：n := FC_DL_DeadtimeTapCalc(tDeadtime := T#2S, tSample := T#100MS,
 *                                       bSaturated => bSat, bValid => bOk);
 * 注意：n = 20；bSaturated = TRUE 时结果为饱和钳位值，禁入 Smith 本体。
 *-----------------------------------------------------------------------------*)
FUNCTION FC_DL_DeadtimeTapCalc : DINT
VAR_INPUT
    tDeadtime : TIME;                  // 死区时间 [毫秒] / Dead time [ms]
    tSample   : TIME;                  // 离散采样拍长 [毫秒] / Discrete sample period [ms]
END_VAR
VAR_OUTPUT
    bSaturated : BOOL;                 // 饱和钳位声明（TRUE 时结果为钳位值）/ Saturation declaration
    bValid     : BOOL;                 // 结果有效标志，FALSE 时返回哨兵 0 / Result validity flag
END_VAR
VAR CONSTANT
    DL_DT_DINTMAX : DINT   := 2147483647; // DINT 正向上限 / DINT positive ceiling
    DL_DT_EPS     : LREAL  := 1.0E-6;   // 余量进位容差 [拍] / Carry tolerance [taps]
    DL_DT_ZERO    : DINT   := 0;        // 无效哨兵返回值 / Sentinel return for invalid
    DL_DT_MS_PER_S: LREAL  := 1000.0;   // 毫秒→秒换算系数 [毫秒每秒] / ms-to-s scale [ms per s]
END_VAR
VAR
    fDeadSec : LREAL;                  // 死区时间换算秒 [秒] / Dead time in seconds [s]
    fSmpSec  : LREAL;                  // 采样拍长换算秒 [秒] / Sample period in seconds [s]
    fQuot    : LREAL;                  // 实数商 [拍] / Real quotient [taps]
    nQuot    : DINT;                   // TRUNC 整商 [拍] / Truncated integer quotient [taps]
    fRemain  : LREAL;                  // 余量 [拍] / Remainder fraction [taps]
END_VAR

// ---- 段 1｜出口默认值（纯函数无实例，无定时器/沿刷新义务）----
bSaturated := FALSE;                  // 饱和声明默认 FALSE / Saturation preset FALSE
bValid := FALSE;                      // 缺省无效 / Invalid by default

// ---- 段 2｜TIME → 秒换算（标准显式转换 R10；TIME 上限 DWORD 毫秒域足够）----
fDeadSec := DINT_TO_LREAL(TIME_TO_DINT(tDeadtime)) / DL_DT_MS_PER_S; // 死区秒值 [秒] / Dead time seconds
fSmpSec  := DINT_TO_LREAL(TIME_TO_DINT(tSample)) / DL_DT_MS_PER_S;   // 拍长秒值 [秒] / Sample seconds

// ---- 段 3｜域闸：拍长正域 + 死区非负域（TIME 为无符号毫秒，仍双闸防御）----
IF (fSmpSec <= 0.0) OR (fDeadSec < 0.0) THEN
    FC_DL_DeadtimeTapCalc := DL_DT_ZERO; // 域外拒绝：哨兵零返回 / Out of domain, refused
    RETURN;                            // 结构早退 / early exit
END_IF

// ---- 段 4｜商主体与取整纪律：先 TRUNC 整商，余量超容差才进位（禁 TRUNC+1）----
fQuot   := fDeadSec / fSmpSec;        // 实数商 [拍]，分母已过正域闸 / Real quotient, denominator gated
IF fQuot <> fQuot THEN                // 商非有限兜底（双有限入参理论上不可达，R90 复检）
    FC_DL_DeadtimeTapCalc := DL_DT_ZERO; // 非有限商哨兵返回 / Non-finite quotient, sentinel return
    RETURN;                            // 结构早退 / early exit
END_IF
IF fQuot >= DINT_TO_LREAL(DL_DT_DINTMAX) THEN // 实数上限兜底：商超 DINT 域直接饱和（防 TRUNC 溢出回绕，R28）
    FC_DL_DeadtimeTapCalc := DL_DT_DINTMAX; // 饱和钳位出口 / Saturating outlet
    bSaturated := TRUE;                // 饱和声明置位 / Saturation declared
    bValid := TRUE;                    // 饱和是合法结论（调用方判 bSaturated）/ Saturation is a valid conclusion
    RETURN;                            // 结构早退 / early exit
END_IF
nQuot   := TRUNC(fQuot);              // TRUNC 整商（向零取整，商恒非负；上限已预闸不溢）/ Truncated quotient, ceiling pre-gated
fRemain := fQuot - DINT_TO_LREAL(nQuot); // 余量 [拍] / Remainder fraction
IF fRemain > DL_DT_EPS THEN           // 余量超容差才进位（纯整除不虚进一位）/ Carry only on real remainder
    IF nQuot >= DL_DT_DINTMAX THEN
        nQuot := DL_DT_DINTMAX;      // 整商已顶上限：饱和钳位不进位（防回绕）/ Quotient at ceiling, saturate
        bSaturated := TRUE;          // 饱和声明置位 / Saturation declared
    ELSE
        nQuot := nQuot + 1;          // 正常进位一位 / Normal one-tap carry
    END_IF
END_IF
FC_DL_DeadtimeTapCalc := nQuot;       // 离散拍数 [拍] / Discrete tap count
bValid := TRUE;                       // 全部防御通过：结果有效 / Result valid
END_FUNCTION

(* ---- FC_DL_DepositionUniformityCalc.st ---- *)
(*
  DL Factory R88 | FC_DL_DepositionUniformityCalc
  功能：由固定五点膜厚算均匀性 (max-min)/(2·mean)×100%，并按 3% 判合格（不用数组，逐点标量入参）
  开源溯源：无（clean-room 自研，依据公开工艺公式 膜厚均匀性式 (max-min)/(2·mean)，许可证=MIT，借鉴点=公式结构）
  规则：R1-R16 全遵守；R88 简单件标量形（纯标量入参出参，无循环体、无方法、无属性、无数组）
*)
FUNCTION FC_DL_DepositionUniformityCalc : REAL
VAR_INPUT
    fT1 : REAL := 100.0; // 测点 1 膜厚（中心） [nm] / thickness at site 1, centre [nm]
    fT2 : REAL := 98.0; // 测点 2 膜厚 [nm] / thickness at site 2 [nm]
    fT3 : REAL := 102.0; // 测点 3 膜厚 [nm] / thickness at site 3 [nm]
    fT4 : REAL := 99.0; // 测点 4 膜厚 [nm] / thickness at site 4 [nm]
    fT5 : REAL := 101.0; // 测点 5 膜厚 [nm] / thickness at site 5 [nm]
    fTolPct : REAL := 3.0; // 均匀性公差上限 [%] / uniformity tolerance [%]
END_VAR
VAR_OUTPUT
    fUniformityPct : REAL; // 膜厚不均匀度 [%] / thickness non uniformity [%]
    xPass : BOOL; // TRUE=不均匀度不超过公差 [-] / TRUE when within tolerance [-]
END_VAR
VAR
    fMaxT : REAL; // 五点最大膜厚 [nm] / maximum thickness [nm]
    fMinT : REAL; // 五点最小膜厚 [nm] / minimum thickness [nm]
    fMeanT : REAL; // 五点平均膜厚（除零判据） [nm] / mean thickness, the divisor [nm]
END_VAR

// 段 1｜出口预置
FC_DL_DepositionUniformityCalc := -1.0; // 哨兵返回 -1（无效） [-] / sentinel return -1, invalid [-]
fUniformityPct := 0.0; // 不均匀度预置零 [%] / non uniformity preset zero [%]
xPass := FALSE; // 合格位预置 FALSE（未判定前不认合格） [-] / pass flag preset false [-]

// 段 2｜非有限拦截 + 域闸
IF NOT (fT1 > -1.0E30 AND fT1 < 1.0E30) OR NOT (fT2 > -1.0E30 AND fT2 < 1.0E30) OR NOT (fT3 > -1.0E30 AND fT3 < 1.0E30) THEN
    RETURN; // 测点 1/2/3 任一非有限即拒算 [-] / any non finite thickness rejected [-]
END_IF
IF NOT (fT4 > -1.0E30 AND fT4 < 1.0E30) OR NOT (fT5 > -1.0E30 AND fT5 < 1.0E30) OR NOT (fTolPct > -1.0E30 AND fTolPct < 1.0E30) THEN
    RETURN; // 测点 4/5 与公差任一非有限则判据静默失效，故先拦 [-] / these pins must be finite [-]
END_IF
IF fT1 < 0.0 OR fT2 < 0.0 OR fT3 < 0.0 OR fT4 < 0.0 OR fT5 < 0.0 THEN
    RETURN; // 膜厚非负闸：负厚度无物理意义 [nm] / non negative thickness gate [nm]
END_IF
IF fTolPct <= 0.0 THEN
    RETURN; // 公差正域闸：非正公差会使判定恒不合格 [%] / positive tolerance gate [%]
END_IF

// 段 3｜计算（五点极值 + 算术平均，等价 max/min/sum 三路归约）
fMaxT := MAX(MAX(fT1, fT2), MAX(fT3, MAX(fT4, fT5))); // 三级取大得 max [nm] / nested maximum [nm]
fMinT := MIN(MIN(fT1, fT2), MIN(fT3, MIN(fT4, fT5))); // 三级取小得 min [nm] / nested minimum [nm]
fMeanT := (fT1 + fT2 + fT3 + fT4 + fT5) * 0.2; // nm × 0.2 = nm，五点算术平均（乘 0.2 替除 5） [nm] / [nm]
IF fMeanT < 1.0E-9 THEN
    RETURN; // 除法前分母闸：平均膜厚必须大于 1E-9（全零测点无意义） [nm] / denominator gate [nm]
END_IF
fUniformityPct := (fMaxT - fMinT) / (2.0 * fMeanT) * 100.0; // (nm ÷ nm) × 100 = %，极差折半归一到均值 [%] / [%]

// 段 4｜判定与饱和
IF NOT (fUniformityPct > -1.0E30 AND fUniformityPct < 1.0E30) THEN
    RETURN; // 结果非有限再拦一次 [-] / re-check the result for finiteness [-]
END_IF
xPass := fUniformityPct <= fTolPct; // 不均匀度不超过公差即合格（含边界） [%] / within tolerance, boundary included [%]

// 段 5｜出口自检
IF fMaxT < fMinT THEN
    RETURN; // 出口自检：极值关系被破坏说明归约链出错 [nm] / extremum order violated [nm]
END_IF
FC_DL_DepositionUniformityCalc := fUniformityPct; // 返回膜厚不均匀度 [%] / return the non uniformity [%]
END_FUNCTION
